(* IEC 61131-3 sources: daoli-st-library/DL_Base (part 13) *)

(* ---- FB_DL_InterlockMatrix.st ---- *)
(*==============================================================================
 * 组件名称 (Component)  : FB_DL_InterlockMatrix
 * 所属子库 (Sublibrary) : DL_Base
 * 当前版本 (Version)    : 1.0.1
 * 兼容性   (Platform)   : CODESYS 3.5 / TwinCAT 3 / 汇川 InoProShop / Machine Expert
 *                         仅依赖 Standard.library（R_TRIG / SHR / SHL），零厂商方言
 * 功能描述 (Function)   : 16 路安全联锁条件的汇总与首因（首出）追踪。
 *                         全部停机级条件满足才给出唯一一个运行许可位 bPermitToRun；
 *                         条件失效的瞬间锁存"第一个失效的通道号 + 完整位图 + 全局序号"，
 *                         复位后若条件仍未恢复，复位挂起而不清锁存。
 *                         解决两类现场顽疾：①停机后十条联锁同时报，维修工不知道先查哪条；
 *                         ②复位键一按就放行，根因被掩盖，第二天同一故障再来一次。
 *                         本块只回答"能不能开机"，"先看哪条报警"由报警管理组件负责。
 *
 * 【取反掩码真值表 / Invert-mask truth table（边界 B7）】
 *   raw  invert  →  有效值   现场含义
 *    0     0     →   0       常开触点未动作，条件不满足
 *    1     0     →   1       常开触点动作，条件满足
 *    0     1     →   1       常闭触点未断开（如未拍下的急停），条件满足
 *    1     1     →   0       常闭触点已断开（急停被拍下），条件不满足
 *   结论：常闭接线的急停、安全门、油压过低开关，必须把对应 invert 位置 1。
 *
 * 【失真与语义披露 / Distortion disclosure】
 *   1) 首因只在"停机级位图由 0 变非 0"的那一拍捕获。若两路在同一扫描周期内失效，
 *      扫描粒度内无法排序，此时取最低索引为代表值、置 bFirstOutSimult，并锁存整张位图；
 *      严禁在 HMI 上编造"谁先谁后"。
 *   2) 提示级失效不参与首因、不阻断许可，避免"料仓低"把停机首因挤掉。
 *   3) 上电首扫即锁存（不等沿）：冷启动时的首因可能只是"本来就断着"的条件，
 *      不代表本次停机原因，bLatchedAtStartup 用于区分这两种情形。
 *
 * 开源溯源 (Origin)     : 原创实现（参考 ISA-18.2 的首出方法论与西门子 LGF 位逻辑功能组的
 *                         参数分类，clean-room 编写，未复制任何源码）
 * 本文件内含       : TYPE  E_DL_InterlockState（配套枚举，归属 DL_Base）
 *                    FB    FB_DL_InterlockMatrix
 * 依赖     (Depends)    : 无 DL_ 内部依赖；Standard.library: R_TRIG / SHR / SHL
 * 红线自检 (Redline)    : R1 ✓ 零全局变量表与外部变量引用 ｜ R2 ✓ 零物理 IO 地址直写
 *                         R3 ✓ 纯 IEC 61131-3（位操作一律 SHR/SHL + AND/OR，无位访问方言）
 *                         R4 ✓ 配置非法即禁放行 + 复位挂起 + 序号饱和 + 索引钳位
 *                         R5 ✓ 全变量中英双语同行注释 ｜ R6 ✓ 五态 ENUM + CASE + ELSE 兜底
 *                         R7 ✓ 边沿实例主体最前部无条件刷新（本块仅一个实例）
 * 修订历史 (Revision)   :
 *   2026-11-14  v1.0.0  首版入库（Phase 1 收口批次 · R3）
 *   2026-11-16  v1.0.1  R13 机检 R39 修复：段 8 未使能覆盖原先把 eStateInt 无条件
 *                       改写为 eDisabled，而 eLatched / eFault 两态的复位沿消化
 *                       位于其后段 9 的 CASE 分支内——禁用期间按下的复位沿被整拍
 *                       吞掉，首因锁存与配置故障均需二次复位才清除。改为两个持有
 *                       复位沿的状态不被禁用覆盖，其余态行为不变
 *============================================================================*)

(*-----------------------------------------------------------------------------
 * 枚举: E_DL_InterlockState（归属 DL_Base，与 FB_DL_InterlockMatrix 同文件）
 * 含义: 联锁矩阵主状态。数值步长留空位便于后续插态而不破坏已有工程。
 *----------------------------------------------------------------------------*)
TYPE E_DL_InterlockState :
(
    eDisabled  := 0,     // 未使能：许可强制 FALSE，锁存内容保持 / Disabled, permit forced FALSE, latches kept
    eBlocked   := 10,    // 条件不满足：许可 FALSE，等待恢复 / Blocked, waiting for the conditions
    ePermitted := 20,    // 全部停机级条件满足，许可 TRUE / Permitted, all trip-class conditions OK
    eLatched   := 30,    // 首因已锁存，等待复位 / First-out latched, waiting for reset
    eFault     := 99     // 配置非法：无任何停机级通道，需改配置后复位 / Invalid configuration
);
END_TYPE

(*==============================================================================
 * 功能块: FB_DL_InterlockMatrix
 * 调用约定: 每个扫描周期无条件调用一次；abConditionOk 必须每拍整体刷新。
 * 无状态泄漏: 全部状态驻留于实例私有 VAR，零全局引用，可多机组并行实例化。
 *============================================================================*)
FUNCTION_BLOCK FB_DL_InterlockMatrix
VAR_INPUT
    abConditionOk : ARRAY[0..15] OF BOOL;     // 16 路原始条件，TRUE = 满足（上限 16 路）/ Raw conditions, TRUE = OK, max 16
    auInvertMask  : WORD := 16#0000;          // 取反掩码，bit=1 表示该路原始信号需取反 / Invert mask, bit=1 inverts that channel
    auTripMask    : WORD := 16#FFFF;          // 停机级掩码，bit=1 = 停机级，bit=0 = 提示级 / Trip-class mask, bit=1 is trip class
    bEnable       : BOOL := TRUE;             // 使能，FALSE 时许可 FALSE 且不清锁存 / Enable, FALSE forces permit down but keeps latches
    bReset        : BOOL;                     // 上升沿：清除首因锁存（条件未恢复则挂起）/ Rising edge: clear the first-out latch
END_VAR
VAR_OUTPUT
    bPermitToRun      : BOOL;                 // 运行许可（唯一放行信号）/ Run permit, the only release signal
    bFirstOutValid    : BOOL;                 // 首因有效 / First-out valid
    nFirstOutIndex    : INT;                  // 首因通道号 0..15，-1 = 无 / First-out channel 0..15, -1 = none
    uFirstOutMask     : WORD;                 // 首因位图（同拍多点时多 bit）/ First-out bitmap, multi-bit on simultaneous trips
    uFirstOutSeq      : UDINT;                // 首因发生的全局序号（单调递增）/ First-out global sequence, monotonic
    bFirstOutSimult   : BOOL;                 // 首因为同拍多点失效，扫描粒度内不可排序 / Simultaneous first-out, unorderable
    bLatchedAtStartup : BOOL;                 // 首因发生在上电首扫（冷启动即不满足）/ Latched during the first scan
    uTripActiveMask   : WORD;                 // 当前失效的停机级通道位图 / Currently failed trip channels
    uWarnActiveMask   : WORD;                 // 当前失效的提示级通道位图 / Currently failed warning channels
    bResetPending     : BOOL;                 // 复位挂起：已按复位但条件未恢复 / Reset pending, conditions not restored
    bError            : BOOL;                 // 故障标志（配置类锁存）/ Fault flag, configuration fault latched
    uErrorId          : UDINT;                // 故障码，0 = 无故障 / Error code, 0 = no error
    eState            : E_DL_InterlockState;  // 当前状态（供 HMI 诊断）/ Current state for HMI diagnosis
END_VAR
VAR
    fbTrigReset     : R_TRIG;                 // 复位上升沿检测实例 / Reset rising edge detector
    auEffOk         : ARRAY[0..15] OF BOOL;   // 取反后的有效条件（上限 16 路）/ Effective conditions after inversion, max 16
    uTripNow        : WORD;                   // 本拍失效的停机级位图 / Failed trip channels this scan
    uWarnNow        : WORD;                   // 本拍失效的提示级位图 / Failed warning channels this scan
    uPrevTripNow    : WORD;                   // 上一拍失效的停机级位图（判沿用）/ Previous trip bitmap, for edge detection
    uLatchMask      : WORD;                   // 锁存的首因位图 / Latched first-out bitmap
    uFirstOutSeqInt : UDINT;                  // 首因序号的内部副本 / Internal copy of the first-out sequence
    uBitMask        : WORD;                   // 单通道取位探针 / Single-channel bit probe
    nLatchIdx       : INT;                    // 锁存的首因通道号，-1 = 无 / Latched first-out index, -1 = none
    nNewLowest      : INT;                    // 本拍首个失效通道（最低索引）/ Lowest failed index this scan
    nBitCount       : INT;                    // 本拍失效通道总数 / Number of failed channels this scan
    nIdx            : INT;                    // 通道遍历索引 / Channel loop index
    uSeqCounter     : UDINT;                  // 全局序号计数器 / Global sequence counter
    eStateInt       : E_DL_InterlockState;    // 主状态机内部当前态 / Internal state of the main state machine
    bInv            : BOOL;                   // 该通道是否取反 / Whether this channel is inverted
    bConfigInvalid  : BOOL;                   // 本拍配置是否非法（无停机级通道）/ Configuration invalid this scan
    bConfigLatch    : BOOL;                   // 配置故障锁存 / Configuration fault latched
    bNewEvent       : BOOL;                   // 本拍出现新的停机级失效事件 / A new trip event started this scan
    bStartupScan    : BOOL := TRUE;           // 上电首扫标志 / First-scan flag
END_VAR
VAR CONSTANT
    DL_ILK_CHANNELS : INT  := 16;             // 通道数，必须等于数组维度 / Channel count, must match the array dimension
    DL_ILK_IDX_NONE : INT  := -1;             // 无效通道号哨兵 / No-channel sentinel
    DL_ILK_BIT0     : WORD := 16#0001;        // 最低位掩码 / Least significant bit mask
    DL_ILK_SEQ_MAX  : UDINT := 16#FFFF_FFFE;  // 序号饱和值 / Sequence saturation value
END_VAR

(*------------------------------------------------------------------------------
 * 段 1｜无条件刷新区（红线 R7）
 *      Unconditional refresh zone, placed at the very top of the body
 *-----------------------------------------------------------------------------*)
fbTrigReset(CLK := bReset);

(*------------------------------------------------------------------------------
 * 段 2｜上电首扫（边界 B2）：索引与位图必须显式置为哨兵值，不能依赖默认零
 *      First-scan init: the index must be forced to the sentinel, never left at zero
 *      0 号通道是合法的首因值，用 0 当"无首因"会让 HMI 永远显示 CH0 故障
 *-----------------------------------------------------------------------------*)
IF bStartupScan THEN
    nLatchIdx    := DL_ILK_IDX_NONE;
    uLatchMask   := 16#0000;
    uPrevTripNow := 16#0000;
    uSeqCounter  := 0;
    eStateInt    := E_DL_InterlockState.eBlocked;
END_IF

(*------------------------------------------------------------------------------
 * 段 3｜有效条件求值（边界 B7）：有效 = 原始 XOR 取反位
 *      Effective value = raw XOR invert, one pass over the 16 channels
 *      真值表见文件头；常闭接线的急停必须置 invert 位，否则"拍下急停"会被判为满足
 *      Normally-closed devices must set the invert bit, otherwise pressing the e-stop
 *      would read as a satisfied condition
 *-----------------------------------------------------------------------------*)
FOR nIdx := 0 TO (DL_ILK_CHANNELS - 1) DO
    uBitMask      := SHR(auInvertMask, nIdx) AND DL_ILK_BIT0;
    bInv          := (uBitMask <> 16#0000);
    auEffOk[nIdx] := abConditionOk[nIdx] XOR bInv;
END_FOR

(*------------------------------------------------------------------------------
 * 段 4｜分类汇总（边界 B6）：停机级进 uTripNow，提示级进 uWarnNow
 *      Classification: trip-class feeds the bitmap, warning-class only reports
 *      位操作一律 SHR/SHL 取位置位，禁止位访问方言，保证三平台同码
 *-----------------------------------------------------------------------------*)
uTripNow := 16#0000;
uWarnNow := 16#0000;

FOR nIdx := 0 TO (DL_ILK_CHANNELS - 1) DO
    IF NOT auEffOk[nIdx] THEN
        uBitMask := SHR(auTripMask, nIdx) AND DL_ILK_BIT0;
        IF uBitMask <> 16#0000 THEN
            uTripNow := uTripNow OR SHL(DL_ILK_BIT0, nIdx);
        ELSE
            uWarnNow := uWarnNow OR SHL(DL_ILK_BIT0, nIdx);
        END_IF
    END_IF
END_FOR

(*------------------------------------------------------------------------------
 * 段 5｜首因定位（边界 B3/B4）：求最低索引与失效总数
 *      First-out localisation: find the lowest failed index and the failed count
 *      同拍多路失效时无法排序，只能给代表值与位图，绝不编造先后
 *-----------------------------------------------------------------------------*)
nNewLowest := DL_ILK_IDX_NONE;
nBitCount  := 0;

FOR nIdx := 0 TO (DL_ILK_CHANNELS - 1) DO
    uBitMask := SHR(uTripNow, nIdx) AND DL_ILK_BIT0;
    IF uBitMask <> 16#0000 THEN
        nBitCount := nBitCount + 1;
        IF nNewLowest < 0 THEN
            nNewLowest := nIdx;
        END_IF
    END_IF
END_FOR

(*------------------------------------------------------------------------------
 * 段 6｜首因捕获：上电首扫特殊处理（边界 B2），其余按 0→非 0 的沿捕获
 *      First-out capture: special case on the first scan, edge-triggered afterwards
 *      锁存后不再被新故障覆盖——首因就是首因，覆盖等于把根因洗掉
 *      Once latched the value is never overwritten: the first cause stays the first cause
 *      首扫时 uPrevTripNow 已被置 0，因此"上电本来就不满足"同样走这条沿路径，
 *      只是序号从 1 开始并被标记为 bLatchedAtStartup
 *-----------------------------------------------------------------------------*)
bNewEvent := FALSE;

IF (uTripNow <> 16#0000) AND (uPrevTripNow = 16#0000) THEN
    bNewEvent := TRUE;
END_IF

IF bNewEvent THEN

    IF uSeqCounter < DL_ILK_SEQ_MAX THEN
        uSeqCounter := uSeqCounter + 1;
    ELSE
        uErrorId := 16#0001_0007;
    END_IF

    IF nLatchIdx < 0 THEN
        nLatchIdx         := nNewLowest;
        uLatchMask        := uTripNow;
        uFirstOutSeqInt   := uSeqCounter;
        bFirstOutSimult   := (nBitCount > 1);
        bLatchedAtStartup := bStartupScan;
    END_IF

END_IF

uPrevTripNow := uTripNow;

(*------------------------------------------------------------------------------
 * 段 7｜配置校验（边界 B1，fail-safe 第一原则）
 *      Configuration check: no trip-class channel means the permit can never be gated
 *      无任何停机级通道时若默认放行，等于把"没配置"当成"全部满足"，这是最危险的缺省
 *      Defaulting to permit when nothing is configured is the most dangerous default
 *-----------------------------------------------------------------------------*)
bConfigInvalid := (auTripMask = 16#0000);

IF bConfigInvalid THEN
    bConfigLatch := TRUE;
END_IF

IF bConfigLatch THEN
    uErrorId  := 16#0002_0004;
    eStateInt := E_DL_InterlockState.eFault;
END_IF

(*------------------------------------------------------------------------------
 * 段 8｜未使能处理：许可撤销、锁存保持（使能不是复位）
 *      Disabled: the permit drops but the latches survive, enabling is not resetting
 *      R39 纪律：复位沿只在发生的那一拍为真，其消化权归段 9 的 eLatched 与 eFault
 *      两个分支所有。本段若无条件把状态改写成 eDisabled，则禁用期间按下的复位沿
 *      在本拍即被抹掉（段 9 走 eDisabled 分支，两处复位判据都摸不到该沿），首因
 *      锁存与配置故障只能靠操作员补按第二次复位——故这两态不参与禁用覆盖。
 *      R39: the reset edge lives for exactly one scan and is consumed inside the CASE
 *      branches of eLatched and eFault, so the disable override must leave both
 *      states untouched; otherwise a reset pressed while disabled is lost and the
 *      first-out latch needs a second press. The other states keep the old behaviour.
 *-----------------------------------------------------------------------------*)
IF (eStateInt <> E_DL_InterlockState.eLatched)
AND (eStateInt <> E_DL_InterlockState.eFault)
AND (NOT bEnable) THEN
    eStateInt := E_DL_InterlockState.eDisabled;
END_IF

(*------------------------------------------------------------------------------
 * 段 9｜主状态机（红线 R6）：ENUM + CASE + ELSE 兜底
 *      Main state machine with the mandatory ELSE fallback
 *-----------------------------------------------------------------------------*)
CASE eStateInt OF

    E_DL_InterlockState.eDisabled:
        IF bEnable THEN
            IF bConfigLatch THEN
                eStateInt := E_DL_InterlockState.eFault;
            ELSE
                eStateInt := E_DL_InterlockState.eBlocked;
            END_IF
        END_IF

    E_DL_InterlockState.eBlocked:
        IF uTripNow <> 16#0000 THEN
            eStateInt := E_DL_InterlockState.eLatched;
        ELSE
            eStateInt := E_DL_InterlockState.ePermitted;
        END_IF

    E_DL_InterlockState.ePermitted:
        (* 任一停机级失效立即降级，许可在同一拍撤销（状态即许可） *)
        (* Any trip-class failure demotes at once, the permit drops in the same scan *)
        IF uTripNow <> 16#0000 THEN
            eStateInt := E_DL_InterlockState.eLatched;
        END_IF

    E_DL_InterlockState.eLatched:
        (* 边界 B5：条件未恢复时复位只挂起、不清锁存 *)
        (* Reset only pends while a trip condition is still present *)
        IF fbTrigReset.Q THEN
            IF uTripNow = 16#0000 THEN
                nLatchIdx         := DL_ILK_IDX_NONE;
                uLatchMask        := 16#0000;
                uFirstOutSeqInt   := 0;
                bFirstOutSimult   := FALSE;
                bLatchedAtStartup := FALSE;
                bResetPending     := FALSE;
                eStateInt         := E_DL_InterlockState.eBlocked;
            ELSE
                bResetPending := TRUE;
            END_IF
        END_IF

    E_DL_InterlockState.eFault:
        (* 配置故障：必须先把停机级掩码改对，再按复位退出 *)
        (* Configuration fault: fix the trip mask first, then reset *)
        IF fbTrigReset.Q AND (NOT bConfigInvalid) THEN
            bConfigLatch := FALSE;
            uErrorId     := 16#0000_0000;
            eStateInt    := E_DL_InterlockState.eBlocked;
        END_IF

    ELSE
        (* 非法状态拦截：不做隐式恢复，直接锁存上报 *)
        (* Illegal state interception: no implicit recovery, latch and report *)
        eStateInt := E_DL_InterlockState.eFault;
        uErrorId  := 16#0001_0005;

END_CASE;

(*------------------------------------------------------------------------------
 * 段 10｜输出单一出口（范式 P-05）
 *      Single output exit: the permit derives from the state exactly once
 *      分支内只改状态，许可位只在此处派生，"多处置位、漏撤一处"从结构上不可能
 *-----------------------------------------------------------------------------*)
bPermitToRun      := (eStateInt = E_DL_InterlockState.ePermitted) AND bEnable AND (NOT bConfigLatch);
bFirstOutValid    := (nLatchIdx >= 0);
nFirstOutIndex    := nLatchIdx;
uFirstOutMask     := uLatchMask;
uFirstOutSeq      := uFirstOutSeqInt;
uTripActiveMask   := uTripNow;
uWarnActiveMask   := uWarnNow;
bError            := (eStateInt = E_DL_InterlockState.eFault) OR bConfigLatch;
eState            := eStateInt;

(* 首扫标志在主体末尾撤销：段 6 需要它区分"冷启动即不满足"与"运行中失效" *)
(* The first-scan flag is cleared only here, stage 6 needs it for the cold-start case *)
bStartupScan := FALSE;
END_FUNCTION_BLOCK

(* ---- FB_DL_LastGoodValueHold.st ---- *)
(*
  ==================================================================
  组件名 Component  : FB_DL_LastGoodValueHold
  分类   Category   : DL_Base
  前缀   Naming     : FB_DL_ ｜ b/n/u/f/t/e 类型前缀制（R265）
  版本   Version    : 1.0.0
  功能   Purpose    : NE43 信号质量失效保持件：bSigOk=TRUE（质量好）时
                      透传 fInVal 并刷新保持载体；bSigOk=FALSE（NE43 超
                      量程/欠量程/断线诊断失效）时输出冻结为最后有效值
                      fLastGood，同时 tonStale 累计陈旧时长，超 tStaleMax
                      置信息码 01 与 bStale（输出仍保持最后有效值，不静
                      默）。失效时无历史有效值（首件语义）bValid=FALSE
                      并置信息码 03。tStaleMax ≤ 0 配置非法电平面码 02。
  来源   Source     : t2-8-ne43（NE43 欠量程/超量程诊断语义为公开行业
                      口径（NAMUR NE43），实现零源码复制）
  互引   Cross-ref  : FB_DL_AnalogOutFailsafe（同族失效安全件：其面向模
                      出通道失效替代，本件面向模拟量输入信号质量保持，
                      二者可级联——本件输出喂其输入）
  平台   Platform   : 纯 IEC 61131-3（TON/LREAL 四则/TIME 比较）
  依赖   Depends    : 仅 Standard.library（TON 属标准件）
  红线   Redline    : R1 零全局/VAR_EXTERNAL/R2 零 %I/%Q/R3 纯 IEC 标准
                      R4 输入非有限闸 + 配置闸显式 + TON 实例段 0 无条件
                      刷新/R5 全变量双语同行注释/R6 配置故障电平面无状
                      态机（CASE 不适用，头注说明）/R7 tonStale 无条件周
                      期调用/R8 阈值常量化
  契约   Contract   : 码 02 配置非法为电平面（当拍复判）：故障拍 bValid=
                      FALSE、fOut 冻结保持、bError=TRUE，恢复即恢复；
                      码 01/03 为信息级不置 bError。信号恢复（bSigOk 上
                      升）即透传刷新载体并清陈旧计时（TON 随 IN=FALSE
                      自清零，R188 自复位语义）。
  错误码 Codes      : 01【信息级】陈旧超限（保持时长超 tStaleMax，输出
                      仍为最后有效值）
                      02【故障级·电平面】tStaleMax ≤ T#0MS 配置非法
                      03【信息级】失效且无保持载体（从未收到有效值，
                      fOut 冻结 0）
  码位反证 Note     : 01/02/03 分立依据（R90）：01 在时效面（载体存在但
                      老化）、02 在配置面、03 在载体面（从未有过）可观测；
                      03 若并入 01，则「等一等会有值」与「永远不会有值」
                      不可区分，故必须分立；02 为故障级置 bError，与
                      01/03 信息级双通道可区分。
  验收   Acceptance : V1 质量好透传 → fOut=fInVal，bValid ｜ V2 失效 →
                      fOut 冻结最后值，bStale=FALSE（未超限）｜ V3 失效
                      超 tStaleMax → 码 01 + bStale ｜ V4 tStaleMax=0 →
                      码 02（电平面）｜ V5 上电即失效 → 码 03，bValid=
                      FALSE ｜ V6 恢复 → 透传 + 陈旧清零
  变更   Revision   : 2026-11-22  v1.0.0  R67 首版（编码阶段批 3 序 3）
  ==================================================================
*)
FUNCTION_BLOCK FB_DL_LastGoodValueHold
VAR_INPUT
    fInVal    : LREAL := 0.0;      // 输入测量值 [工程单位] / the input measured value
    bSigOk    : BOOL := FALSE;     // 信号质量好（NE43 诊断有效）[-] / the signal quality ok flag
    tStaleMax : TIME := T#60S;     // 陈旧时长上限 [ms]，须 > 0 / the staleness limit, must be positive
END_VAR
VAR_OUTPUT
    fOut     : LREAL := 0.0;       // 保持输出（最后有效值或透传）[工程单位] / the hold output
    bStale   : BOOL := FALSE;      // 陈旧超限指示（码 01 同源）[-] / the stale limit indicator
    bValid   : BOOL := FALSE;      // 输出可用标志（有有效载体且配置合法）[-] / the output usability flag
    bError   : BOOL := FALSE;      // 配置故障标志（电平面，恢复即清，R45 配对）/ the configuration fault flag
    uErrorId : UDINT := 16#0000_0000; // 错误码，0=正常，01/02/03 见头注 [码] / the error code [code]
END_VAR
VAR
    tonStale   : TON;              // 陈旧计时实例，段 0 无条件刷新 / the staleness timer instance refreshed unconditionally
    _fLastGood : LREAL := 0.0;     // 最后有效值保持载体 [工程单位] / the last good value hold carrier
    _bHasLast  : BOOL := FALSE;    // 保持载体是否存在（首件判据）[-] / the carrier existence flag
    _bCfgOk    : BOOL := FALSE;    // 本拍配置有效性 [-] / the per scan configuration validity
    _bSigFin   : BOOL := FALSE;    // 本拍输入有限性 [-] / the per scan input finiteness
END_VAR
VAR CONSTANT
    LGV_FIN_MAX  : LREAL := 1.7976931348623157E308; // LREAL 有限上限 / the finite LREAL limit
    LGV_ERR_NONE : UDINT := 16#0000_0000;           // 无错误 [码] / no error [code]
    LGV_ERR_STALE: UDINT := 16#0000_0001;           // 码 01：陈旧超限（信息级）/ code 01, stale limit, info level
    LGV_ERR_CFG  : UDINT := 16#0000_0002;           // 码 02：配置非法 / code 02, illegal configuration
    LGV_ERR_NOVAL: UDINT := 16#0000_0003;           // 码 03：无保持载体（信息级）/ code 03, no carrier, info level
END_VAR

(*------------------------------------------------------------------------------
 * 段 0｜定时器无条件刷新区（红线 R7）：严禁移入 IF / CASE
 *      The timer instance refreshes unconditionally, never inside a branch
 *-----------------------------------------------------------------------------*)
tonStale(IN := (NOT bSigOk) AND _bHasLast, PT := tStaleMax);  // 陈旧计时（失效且有载体才计时；恢复随 IN=FALSE 自清零，R188）/ the staleness timing, self clearing on recovery

(*------------------------------------------------------------------------------
 * 段 1｜错误码本拍预置 / segment 1, the error code per scan preset
 *-----------------------------------------------------------------------------*)
uErrorId := LGV_ERR_NONE;      // 预置无错误 / preset no error
bStale := FALSE;               // 陈旧指示预清（码 01 同源重算）/ preset the stale indicator

(*------------------------------------------------------------------------------
 * 段 2｜配置闸（电平面，当拍复判，码 02）+ 输入有限性闸
 *      The configuration gate and the input finiteness gate
 *-----------------------------------------------------------------------------*)
_bCfgOk := (tStaleMax > T#0MS);  // 配置闸（TIME 直接比较，三平台一致）/ the configuration gate
_bSigFin := (fInVal = fInVal) AND (ABS(fInVal) <= LGV_FIN_MAX);  // 输入非有限闸（NaN 自反判 + Inf 兜底）/ the input finite gate
IF NOT _bCfgOk THEN
    bError := TRUE;              // 故障标志（R45 配对）/ the fault flag
    uErrorId := LGV_ERR_CFG;     // 码 02 / code 02
    bValid := FALSE;             // 配置非法不出数 / no output on illegal configuration
    RETURN;                      // fOut 冻结保持（头注契约）/ the output frozen
ELSE
    bError := FALSE;             // 配置恢复即清（电平面契约）/ cleared when the configuration recovers
END_IF

(*------------------------------------------------------------------------------
 * 段 3｜质量好相：透传刷新载体（含非有限拒收，码 03 语义延用）
 *      The good quality phase, pass through and refresh the carrier
 *-----------------------------------------------------------------------------*)
IF bSigOk AND _bSigFin THEN
    _fLastGood := fInVal;        // 载体刷新 / refresh the carrier
    _bHasLast := TRUE;           // 载体存在 / the carrier exists
END_IF

(*------------------------------------------------------------------------------
 * 段 4｜失效相与出口映射：透传或保持，码 01/03 信息级
 *      The failed phase and the outlet mapping, the info codes
 *-----------------------------------------------------------------------------*)
IF bSigOk AND _bSigFin THEN
    fOut := fInVal;              // 透传 / pass through
ELSIF _bHasLast THEN
    fOut := _fLastGood;          // 保持最后有效值（锁存载体，非实时镜像混用）/ hold the last good value, the carrier not a live mirror
ELSE
    fOut := 0.0;                 // 无载体冻结 0（头注契约）/ frozen zero without a carrier
END_IF
IF (NOT bSigOk) OR (NOT _bSigFin) THEN
    IF NOT _bHasLast THEN
        uErrorId := LGV_ERR_NOVAL;  // 码 03：失效且从未有载体（信息级）/ code 03, no carrier, info level
        bValid := FALSE;            // 无值可保 / nothing to hold
    ELSE
        IF tonStale.Q THEN
            uErrorId := LGV_ERR_STALE;  // 码 01：陈旧超限（信息级，不置 bError）/ code 01, stale, info level
            bStale := TRUE;             // 陈旧指示（与码 01 同源，R191 名实双出口）/ the stale indicator
        END_IF
        bValid := TRUE;             // 有载体即可用（保持值有效语义）/ usable with a carrier
    END_IF
ELSE
    bValid := TRUE;                 // 质量好透传可用 / usable while passing through
END_IF
END_FUNCTION_BLOCK

(* ---- FB_DL_LongPressButton.st ---- *)
(*
  ==================================================================
  组件名 Component  : FB_DL_LongPressButton
  分类   Category   : DL_Base
  前缀   Naming     : FB_DL_ ｜ b/n/u/f/t/e/st 类型前缀制（R265）
  复杂度 Complexity  : 中
  版本   Version    : 1.0.0
  功能   Purpose    : 单按钮短按/长按/超长按三档时序分档（三窗 TON 阈值单拍分档）。
  来源   Source     : self-std（IEC 人机交互时序语义自研）
  平台   Platform   : 纯 IEC 61131-3（Standard.library: TON / R_TRIG / F_TRIG），无私有库
  分工声明 Split     : 与 FB_DL_ToggleButtonBank（模式解算属主）分工——后者做
                      按压次数模式解算；本件做单按钮按持续时长的三档分档
                      （R216 双向互引）。
  作者   Author     : 道莅代码库 · PLC 编程专家（R61）
  归属 Ownership     : 本件无 TYPE 声明；引用件类型全部 IEC 标准原生。
  ------------------------------------------------------------------
  边界 Boundary     :
                      一 三档窗组态闸（R239）：tShort < tLong < tXLong 且三者 > 0，
                         违反判组态非法故障码并冻结分档输出（锁存至复位沿）；
                      二 三窗职责与配比约束（R100）：tonShort < tonLong < tonXLong
                         由组态闸结构性保证；长按/超长按在按压持续中经阈值沿
                         单拍分档，短按在释放沿回判；
                      三 TON / R_TRIG / F_TRIG 全部段 0 无条件周期刷新（禁入分支）；
                      四 三档脉冲为单拍输出，段 1 统一预置 FALSE、分支只写 TRUE
                         （R256），内部 _b* 两段式映射（R187）；
                      五 故障态语义为「冻结保持全假输出」（R191 声明行）；
                      六 故障解除路径：复位沿清锁存（bReset 恒可达，R152 自证）；
                      七 无全局、无外部变量、无物理地址。
  错误码   Codes    :
    16#0001_0640【故障级】三档窗组态非法（tShort < tLong < tXLong 违反或 ≤0），锁存至复位沿
  验收   Acceptance :
    算法已证（脚本）：未跑 ｜ 编译器已证（三平台）：未跑
    V1 按下 200ms 释放（tShort=100/tLong=800/tXLong=2000）→ bShortPress 单拍
    V2 按住 1s → 长按阈值拍 bLongPress 单拍；V3 按住 2.5s → bXLongPress 单拍
    V4 tShort = tLong → 码 0640、三脉冲恒假、锁存待复位
  修订记录 Revision  :
    2026-11-21  v1.0.0  R61 首版（批 2 · 序号 8）
  ==================================================================
*)
FUNCTION_BLOCK FB_DL_LongPressButton
VAR_INPUT
    bBtn   : BOOL := FALSE; // 按钮输入电平 [-] / the button input level
    bReset : BOOL := FALSE; // 故障复位电平，上升沿清锁存 [-] / the fault reset level
    tShort : TIME := T#100MS; // 短按下限阈值 [毫秒]，须 < tLong / the short press lower threshold
    tLong  : TIME := T#800MS; // 长按阈值 [毫秒]，须 < tXLong / the long press threshold
    tXLong : TIME := T#2S;    // 超长按阈值 [毫秒] / the extra long press threshold
END_VAR
VAR_OUTPUT
    bShortPress : BOOL := FALSE; // 短按单拍脉冲（释放沿回判）[-] / the short press one shot
    bLongPress  : BOOL := FALSE; // 长按单拍脉冲（tLong 阈值沿）[-] / the long press one shot
    bXLongPress : BOOL := FALSE; // 超长按单拍脉冲（tXLong 阈值沿）[-] / the extra long press one shot
    bFaulted    : BOOL := FALSE; // 组态故障锁存指示 [-] / the latched configuration fault indicator
    eErr        : UDINT := 16#0000_0000; // 错误码，0 = 正常 / the error code, zero is ok
    bError      : BOOL := FALSE; // 故障锁存位（与锁存同源，R191）/ the fault bit from the same latch
END_VAR
VAR
    _bInit      : BOOL := FALSE; // 首拍初始化标志（R310）/ the first scan flag
    _bFault     : BOOL := FALSE; // 组态故障锁存副本（仅复位沿清除）/ the fault latch copy
    _bShort     : BOOL := FALSE; // 短拍内部位，段 1 预清段 5 映射 / the internal short bit
    _bLong      : BOOL := FALSE; // 长拍内部位 / the internal long bit
    _bXLong     : BOOL := FALSE; // 超长拍内部位 / the internal extra long bit
    _bLongFired : BOOL := FALSE; // 长按已发标记（释放沿判短按排除用，按压期间保持）/ the long fired flag held during the press
    _bXFired    : BOOL := FALSE; // 超长按已发标记 / the extra long fired flag
    _bCfgBad    : BOOL := FALSE; // 组态非法标记（逐拍重算）/ the configuration fault flag recomputed
    rtBtn       : R_TRIG;  // 按钮按下沿实例，段 0 无条件刷新 / the press edge instance
    ftBtn       : F_TRIG;  // 按钮释放沿实例，段 0 无条件刷新 / the release edge instance
    rtReset     : R_TRIG;  // 复位沿实例，段 0 无条件刷新 / the reset edge instance
    rtLongQ     : R_TRIG;  // 长窗到时沿实例，段 0 无条件刷新 / the long window expiry edge instance
    rtXLongQ    : R_TRIG;  // 超长窗到时沿实例，段 0 无条件刷新 / the extra long expiry edge instance
    tonShort    : TON;     // 短窗计时，段 0 无条件刷新 / the short window timer
    tonLong     : TON;     // 长窗计时 / the long window timer
    tonXLong    : TON;     // 超长窗计时 / the extra long window timer
END_VAR

// 段 0｜定时器与沿检测无条件周期刷新（禁入分支，R7）/ segment 0, the unconditional refresh
rtBtn(CLK := bBtn); // 按下沿 / the press edge
ftBtn(CLK := bBtn); // 释放沿 / the release edge
rtReset(CLK := bReset); // 复位沿 / the reset edge
tonShort(IN := bBtn, PT := tShort); // 短窗计时（按压电平驱动）/ the short window timing
tonLong(IN := bBtn, PT := tLong); // 长窗计时 / the long window timing
tonXLong(IN := bBtn, PT := tXLong); // 超长窗计时 / the extra long window timing
rtLongQ(CLK := tonLong.Q); // 长窗到时沿 / the long expiry edge
rtXLongQ(CLK := tonXLong.Q); // 超长窗到时沿 / the extra long expiry edge

// 段 1｜首拍初始化与单拍标志预清（仅单拍标志入清单，FB32-1；R256）/ segment 1, the first scan init and the one shot preset
IF NOT _bInit THEN // 首拍一拍 / the first scan
    _bInit := TRUE; // 置首拍标志 / raise the first scan flag
    _bFault := FALSE; // 故障锁存显式清零 / clear the fault latch explicitly
    _bLongFired := FALSE; // 长发标记显式清零 / clear the long fired flag explicitly
    _bXFired := FALSE; // 超长发标记显式清零 / clear the extra long fired flag explicitly
END_IF
IF rtReset.Q THEN // 复位沿：清故障锁存（解除路径：复位沿恒可达，R152 自证）/ the reset edge clears the latch
    _bFault := FALSE; // 清锁存 / clear the latch
END_IF
_bShort := FALSE; // 短拍预清零 / preset the short bit false
_bLong := FALSE; // 长拍预清零 / preset the long bit false
_bXLong := FALSE; // 超长拍预清零 / preset the extra long bit false
_bCfgBad := FALSE; // 组态标记预清零 / preset the configuration flag false

// 段 2｜组态域闸（三窗严格递增 + 正值，R239，边界一）/ segment 2, the configuration gate
IF (tShort <= T#0S) OR (tLong <= tShort) OR (tXLong <= tLong) THEN // 递增配比违反或非正 / the monotone ratio violated
    _bCfgBad := TRUE; // 置组态非法标记 / raise the configuration flag
    _bFault := TRUE; // 锁存故障（段 5 出口回放）/ latch the fault
END_IF

// 段 3｜按压中阈值沿分档（故障冻结，边界五；沿只在合法态消费）/ segment 3, the threshold edges during the press
IF (NOT _bFault) AND bBtn THEN // 合法态且按压中 / legal and pressed
    IF rtLongQ.Q AND (NOT _bLongFired) AND (NOT _bXFired) THEN // 长窗到时沿首现 / the long expiry edge first seen
        _bLong := TRUE; // 置长拍 / raise the long bit
        _bLongFired := TRUE; // 锁长发标记（释放沿判短按排除）/ latch the long fired flag
    END_IF
    IF rtXLongQ.Q AND (NOT _bXFired) THEN // 超长窗到时沿首现 / the extra long expiry edge first seen
        _bXLong := TRUE; // 置超长拍 / raise the extra long bit
        _bXFired := TRUE; // 锁超长发标记 / latch the extra long fired flag
    END_IF
END_IF

// 段 4｜释放沿回判短按（短按 = 释放时短窗已到而长按未发，边界二）/ segment 4, the release edge judges the short press
IF ftBtn.Q AND (NOT _bFault) THEN // 合法态释放沿 / a legal release edge
    IF tonShort.Q AND (NOT _bLongFired) AND (NOT _bXFired) THEN // 短窗已到且未触发高档 / the short window met with no higher grade fired
        _bShort := TRUE; // 置短拍 / raise the short bit
    END_IF
    _bLongFired := FALSE; // 释放清长发标记（下一按压新起点）/ clear the long fired flag at the release
    _bXFired := FALSE; // 释放清超长发标记 / clear the extra long fired flag
END_IF

// 段 5｜统一出口（内部副本单点映射；故障冻结全假，R191）/ segment 5, the unified outlet with the frozen fault
bShortPress := _bShort AND (NOT _bFault); // 短拍出口 / the short outlet
bLongPress := _bLong AND (NOT _bFault); // 长拍出口 / the long outlet
bXLongPress := _bXLong AND (NOT _bFault); // 超长拍出口 / the extra long outlet
bFaulted := _bFault; // 故障指示出口 / the fault indicator outlet
bError := _bFault; // 故障位出口（与锁存同源，R191）/ the fault bit outlet
IF _bFault THEN // 故障锁存回放（R187）/ the latched fault replays
    eErr := 16#0001_0640; // 故障级：三档窗组态非法 / fault grade, the illegal window configuration
ELSE // 无故障 / no fault
    eErr := 16#0000_0000; // 正常 / ok
END_IF
END_FUNCTION_BLOCK

(* ---- FB_DL_ManualOverride.st ---- *)
(*
  道莅工业代码库 | DL_Base | FB_DL_ManualOverride
  版本: 1.0.0 | 日期: 2026-11-23 | 轮次: R75
  开源溯源: brOscatLib (github.com/brOscatLib) / MIT / 借鉴 MANUAL 覆写的语义，代码为 clean-room 重写
  功能: 手动强制覆写——覆写请求上升沿激活后输出切手动值，最长保持 tMaxHold
        （T#0S = 无限时）超时自动回落自动值；释放沿/禁止输入即时回落；
        激活单拍提示脉冲与超时回落信息码。
  兼容性: CODESYS 3.5 / TwinCAT 3 / 汇川 InoProShop；仅依赖标准 TON / R_TRIG / SEL，零厂商私有库
  接口: 输入 bOverrideReq（沿）/bRelease（沿）/fAutoVal/fManualVal/tMaxHold/
        bInhibit/bReset；输出 bOverride/bOut/bActPulse/bTimedOut/eState/eInfo/nErrId。
  码表: 16#0001_04BC 信息级：覆写超时自动回落（锁存至复位沿）
        16#0001_04BD 信息级：覆写请求被禁止拒绝（当拍重算）
        16#0001_04BE 信息级：覆写中手动值非有限（输出保持最后有效值，当拍重算）
        码段说明：0001 段信息子带 04xx，槽位经全库实扫空闲。
  边界: ① 手动值 NaN 拒绝激活（待机相判码），覆写中手动值变 NaN → 输出保持
        最后有效值并置信息码（冻结语义不穿透坏值）；
        ② bInhibit 在覆写中即时回落自动值（禁止优先于覆写，安全侧）；
        ③ 超时判定仅当 tMaxHold > T#0S 生效（T#0S = 无限保持）；
        ④ TON/R_TRIG 段 0 无条件周期刷新；⑤ 本件全部事件均为信息级，无故障级码；
        ⑥ 零全局耦合。
  邻件比对: ToleranceWindow（单容差窗）与本件无语义交集；S04 E_DL_ControlModeSel
            为本件模式语义配套枚举（后续入库）。
  修订历史: 2026-11-23 v1.0.0 R75 首版（复杂件批 B3 · C11）
*)

TYPE E_DL_MovState :
(
    eIdle    := 0,   // 覆写未激活（输出自动值） | Override inactive, output auto value
    eActive  := 10   // 覆写激活（输出手动值） | Override active, output manual value
);
END_TYPE

TYPE E_DL_MovInfo :
(
    eNone      := 0,  // 无事件 | No event
    eTimeout   := 1,  // 超时自动回落（锁存至复位沿） | Timed out, auto fallback latched
    eInhibit   := 2,  // 请求被禁止拒绝（当拍重算） | Request rejected by inhibit
    eNonFinite := 3   // 手动值非有限（当拍重算，输出保持） | Manual value non-finite, output held
);
END_TYPE

FUNCTION_BLOCK FB_DL_ManualOverride
VAR_INPUT
    bOverrideReq : BOOL := FALSE;   // 覆写请求（上升沿激活）[-] | Override request, rising edge activates
    bRelease     : BOOL := FALSE;   // 释放请求（上升沿回落）[-] | Release request, rising edge falls back
    fAutoVal     : REAL := 0.0;     // 自动值 [工程单位] | Auto value
    fManualVal   : REAL := 0.0;     // 手动值（覆写目标）[工程单位] | Manual value, override target
    tMaxHold     : TIME := T#30S;   // 最长覆写保持，T#0S = 无限 | Max hold duration, T#0S = unlimited
    bInhibit     : BOOL := FALSE;   // 覆写禁止（电平，覆写中即时回落）[-] | Override inhibit level
    bReset       : BOOL := FALSE;   // 复位命令，上升沿清超时锁存 [-] | Reset command, rising edge
END_VAR
VAR_OUTPUT
    bOverride : BOOL;               // 覆写激活态 [-] | Override active state
    fOut      : REAL;               // 选择输出（自动/手动/保持值）[工程单位] | Selected output value
    bActPulse : BOOL;               // 激活单拍提示脉冲 [-] | Activation one-shot pulse
    bTimedOut : BOOL;               // 超时回落锁存标志 [-] | Timed-out latch flag
    eState    : E_DL_MovState;      // 状态出口 | State outlet
    eInfo     : E_DL_MovInfo;       // 事件成因出口 | Event cause outlet
    nErrId    : UDINT;              // 事件码，0 = 无事件 | Event code, 0 = none
END_VAR
VAR
    _eState    : E_DL_MovState := E_DL_MovState.eIdle;   // 内部状态（CASE 唯一写入目标） | Internal state
    _eInfo     : E_DL_MovInfo := E_DL_MovInfo.eNone;     // 事件成因锁存（超时级） | Latched event cause
    _bOverride : BOOL;          // 覆写激活锁存位 | Override active latch bit
    _bTimedOut : BOOL;          // 超时回落锁存位 | Timed-out latch bit
    _bHold     : BOOL;          // 输出保持当拍量（手动值非有限）[-] | Output hold this scan
    _fOutLast  : REAL := 0.0;   // 最后有效输出保持值 [工程单位] | Last valid output hold value
    _bNonFin   : BOOL;          // 手动值非有限当拍量 [-] | Manual value non-finite this scan
    _uInfo     : UDINT;         // 信息码每拍重算 | Info code per scan
    rtReq      : R_TRIG;        // 覆写请求沿实例，段 0 无条件刷新 | Override request edge instance
    rtRel      : R_TRIG;        // 释放沿实例，段 0 无条件刷新 | Release edge instance
    rtReset    : R_TRIG;        // 复位沿实例，段 0 无条件刷新 | Reset edge instance
    rtAct      : R_TRIG;        // 激活沿实例（单拍提示），段 0 无条件刷新 | Activation edge instance for one-shot
    tonHold    : TON;           // 覆写保持计时，段 0 无条件刷新 | Override hold timer
END_VAR

(* —— 段 0：当拍量派生 + 定时器与沿实例无条件周期刷新（R7 红线） —— *)
_bNonFin := (fManualVal <> fManualVal);                                     // 手动值 NaN 自反判 / Manual value NaN self-reflex check
rtReq(CLK := bOverrideReq);                                                 // 请求沿每拍必调 / Request edge every scan
rtRel(CLK := bRelease);                                                     // 释放沿每拍必调 / Release edge every scan
rtReset(CLK := bReset);                                                     // 复位沿每拍必调 / Reset edge every scan
rtAct(CLK := _bOverride);                                                   // 激活态沿（单拍提示用）每拍必调 / Activation edge for one-shot
tonHold(IN := (_eState = E_DL_MovState.eActive) AND (tMaxHold > T#0S), PT := tMaxHold);  // 保持计时，IN 挂激活 ∧ 有限时限 / Hold timer gated by active and finite limit

(* —— 段 1：复位沿清超时锁存 —— *)
IF rtReset.Q THEN
    _bTimedOut := FALSE;                                                    // 清超时锁存位 / Clear timed-out latch
    _eInfo := E_DL_MovInfo.eNone;                                           // 清成因锁存 / Clear latched cause
END_IF

(* —— 段 2：状态机（ENUM + CASE，ELSE 兜底） —— *)
CASE _eState OF

E_DL_MovState.eIdle:
    IF rtReq.Q AND bInhibit THEN
        _uInfo := 16#0001_04BD;                                             // 信息级：请求被禁止拒绝 / Info: request rejected by inhibit
    ELSIF rtReq.Q AND _bNonFin THEN
        _uInfo := 16#0001_04BE;                                             // 信息级：手动值非有限拒绝激活 / Info: non-finite manual refused
    ELSIF rtReq.Q THEN
        _bOverride := TRUE;                                                 // 激活覆写锁存 / Activate override latch
        _eState := E_DL_MovState.eActive;                                   // 进入激活相 / Enter active phase
    END_IF

E_DL_MovState.eActive:
    IF rtRel.Q THEN
        _bOverride := FALSE;                                                // 释放沿回落 / Release edge falls back
        _eState := E_DL_MovState.eIdle;
    ELSIF bInhibit THEN
        _bOverride := FALSE;                                                // 禁止输入即时回落（安全侧优先，边界②）/ Inhibit forces fallback
        _eState := E_DL_MovState.eIdle;
    ELSIF tonHold.Q THEN
        _bOverride := FALSE;                                                // 超时回落 / Timed out, fall back
        _bTimedOut := TRUE;                                                 // 超时锁存（复位沿清）/ Latch timeout
        _eInfo := E_DL_MovInfo.eTimeout;                                    // 归因超时 / Cause: timeout
        _eState := E_DL_MovState.eIdle;
    END_IF

ELSE
    _eState := E_DL_MovState.eIdle;                                         // 非法状态兜底（R6，回落安全侧）/ Illegal state fallback to safe side
    _bOverride := FALSE;                                                    // 非法态覆写强制撤 / Override forced off

END_CASE

(* —— 段 3：出口单点映射（名实同源；选择 + 保持 + 锁存码回放） —— *)
IF _bOverride AND _bNonFin THEN
    _bHold := TRUE;                                                         // 覆写中手动值变坏：保持当拍置位（边界①）/ Manual went bad while active, hold
    _uInfo := 16#0001_04BE;                                                 // 信息级：手动值非有限 / Info: manual non-finite
ELSE
    _bHold := FALSE;                                                        // 正常拍不保持 / No hold on normal scan
END_IF
IF (NOT _bHold) AND (NOT (_bOverride AND _bNonFin)) THEN
    _fOutLast := fManualVal;                                                // 有效拍刷新保持值（手动值载体）/ Refresh hold value on valid manual
END_IF
bOverride := _bOverride;                                                    // 覆写态镜像 / Override mirror
IF _bOverride AND _bNonFin THEN
    fOut := _fOutLast;                                                      // 坏值拍输出保持值（冻结语义）/ Bad-value scan outputs held value
ELSIF _bOverride THEN
    fOut := fManualVal;                                                     // 覆写输出手动值 / Override outputs manual value
ELSE
    fOut := fAutoVal;                                                       // 未覆写输出自动值 / Idle outputs auto value
END_IF
bActPulse := rtAct.Q;                                                       // 激活单拍提示（R_TRIG 单拍化） / Activation one-shot
bTimedOut := _bTimedOut;                                                    // 超时锁存镜像 / Timeout latch mirror
eState := _eState;                                                          // 状态出口 / State outlet
eInfo := _eInfo;                                                            // 成因出口 / Cause outlet
IF _bTimedOut THEN
    nErrId := 16#0001_04BC;                                                 // 超时回落锁存码回放（最高优先）/ Replay timeout code
ELSIF _uInfo <> 16#0000_0000 THEN
    nErrId := _uInfo;                                                       // 当拍信息码 / Per-scan info code
ELSE
    nErrId := 16#0000_0000;                                                 // 无事件 / No event
END_IF

END_FUNCTION_BLOCK

(* ---- FB_DL_MinOnOffGuard.st ---- *)
(*
    组件名称 : FB_DL_MinOnOffGuard
    所属子库 : DL_Base
    当前版本 : 1.0.0
    兼 容 性 : CODESYS V3.5+ / TwinCAT 3 / 汇川 InoProShop；仅依赖 Standard.library
    功能描述 : 最短运行 / 最短停止双守卫，防压缩机、热泵、泵轮值与冷水机组频繁启停的公共原子。
              取舍 ①：用「输出实际在 TRUE 期间的累计时长」判最短运行，而不是「进入某状态后重新计时」——
              若定时器只在 eStarting 与 eHolding 里跑，请求在 eRunning 撤掉后会重新起算整段 tMinOn，
              实际运行时长翻倍，压缩机照样被拖坏。本件把 eRunning 一并纳入定时器 IN，
              于是 fbMinOn.Q 的语义严格等于「输出已持续 TRUE 达到 tMinOn」。
              取舍 ②：eIdle 的启动条件只看 bReq，不再二次判 fbMinOff.Q —— 若 eIdle 还要等最短停止完成位，
              而该定时器只在 eCooldown 里通电，则 Q 在 eIdle 恒为 FALSE，状态机将永远起不来（本件修正了这个死锁形态）。
              最短停止由「必须走完 eCooldown 才回 eIdle」保证，语义不减。
              取舍 ③：参数非法不停机 —— 守卫时间填成负值属于参数错误，钳零后继续跑并发故障码；
              让一条产线因为一个 HMI 输入框的负号而停机，代价远大于收益。
              取舍 ④：bEnable = FALSE 走安全侧 —— 立即输出 FALSE 并回 eIdle，忽略最短运行；
              安全优先于设备寿命，两者冲突时永远选安全。
    开源溯源 : 原创实现（T0-2 变体线）。ROADMAP 中「防频繁启停」四条待办的公共原子，无外部源码参考，；本件为 IEC 61131-3 标准语义的道莅防御性实现（原创实现，零外部源码复制）。
              状态机、码位、钳位策略 100% 自有。
    本文件内含 : FUNCTION_BLOCK FB_DL_MinOnOffGuard
                 同文件 TYPE E_DL_MinOnOffState（归属本子库，全库唯一）
    依 赖 : 无 DL_ 内部依赖；Standard.library: TON / R_TRIG
    红线自检 : R1 ✓ 零全局变量与外部变量 ｜ R2 ✓ 零物理 IO 地址
              R3 ✓ 纯 IEC 61131-3 ｜ R4 ✓ 参数钳位 + 非法时间闸 + 非法状态 ELSE 兜底 + 复位沿优先
              R5 ✓ 全变量中英双语同行注释 ｜ R6 ✓ ENUM + CASE + ELSE 兜底（非法状态落 039A 并回安全态）
              R7 ✓ TON / R_TRIG 实例在主体最前部无条件刷新，位于任何 IF 与 CASE 之外
              R8 ✓ 时间上限、零时长、错误码全常量化
    错误码   : 16#0001_0452 [信息级] 时间参数超 24h 已钳上限，bError = FALSE
               16#0001_0453 [信息级] 停机请求被最短运行推迟（进入 eHolding），bError = FALSE
               16#0001_0399 [故障级] 时间参数为负已钳零，不停机，bError = TRUE
               16#0001_039A [故障级] 非法状态（枚举被改写），强制回 eFault 且 bOut = FALSE
               16#0001_039B [故障级] 预留禁用（不得挪用）
    码位总账 : 16#0001_0452 用 / 16#0001_0453 用 ｜ 16#0001_0399 用 / 16#0001_039A 用 / 16#0001_039B 预留
              说明：「启动请求被最短停止阻延」不设独立码 —— 该场景由 eState = eCooldown、bHoldOff 与 tRemaining
              三个输出直接可观测，加强加码属凑槽（R90）。
    遗留假设 : ① TIME 比较与减法按 32 位有符号毫秒口径，加减不越 24h 上限（已由钳位保证），
              故无 TIME 回绕路径；该推导未在三平台逐一实测。
              ② bReset 只在 eFault 内被消费（复位沿实例仍在主体最前部刷新），保证复位沿不被 CASE 前置写吞掉。
    修订历史 :
        2026-11-16  v1.0.0  首版，R21 批次 4 入库
*)

(*-----------------------------------------------------------------------------
 * 枚举: E_DL_MinOnOffState（归属本功能块，与其同文件发布，全库唯一）
 * 含义: 双守卫状态机的六个状态，成员值写死便于工程持久化与在线诊断
 *----------------------------------------------------------------------------*)
TYPE E_DL_MinOnOffState :
(
    eIdle     := 0,     // 空闲：输出 FALSE，最短停止已满，可随时启动 / idle, output low and the minimum off time is satisfied
    eStarting := 10,    // 启动中：输出 TRUE，最短运行计时中 / starting, output high and the minimum on time is counting
    eRunning  := 20,    // 运行中：输出 TRUE，最短运行已满 / running, the minimum on time is satisfied
    eHolding  := 30,    // 保持中：请求已撤但最短运行未满，强制输出 TRUE / holding, the request is gone but the minimum on time is not yet met
    eCooldown := 40,    // 冷却中：输出 FALSE，最短停止计时中 / cooling down, output low and the minimum off time is counting
    eFault    := 99     // 故障锁定：输出 FALSE，需 bReset 上升沿退出 / fault latched, cleared by the rising edge of bReset
);
END_TYPE

FUNCTION_BLOCK FB_DL_MinOnOffGuard
VAR_INPUT
    bEnable         : BOOL := TRUE;      // 使能，FALSE 立即回安全态并忽略最短运行 / enable, FALSE forces the safe state and ignores the minimum on time
    bReq            : BOOL;              // 上层运行请求，TRUE 表示希望设备运行 / run request from the upper layer
    tMinOn          : TIME := T#10S;     // 最短运行时间，负值钳零、超 24h 钳上限 [ms] / minimum on time, clamped at both ends [ms]
    tMinOff         : TIME := T#10S;     // 最短停止时间，负值钳零、超 24h 钳上限 [ms] / minimum off time, clamped at both ends [ms]
    bReset          : BOOL;              // 上升沿清故障并回空闲 / rising edge clears the fault and returns to idle
END_VAR
VAR_OUTPUT
    bOut            : BOOL;              // 实际输出，最终的启停指令 / effective output, the final run command
    bHoldOn         : BOOL;              // TRUE = 正在强制延长运行（停机请求被推迟）/ TRUE while the run time is being extended
    bHoldOff        : BOOL;              // TRUE = 正在强制延长停止（启动请求被阻延）/ TRUE while the stop time is being extended
    tRemaining      : TIME;              // 当前守卫的剩余时间，无守卫时为 0 [ms] / remaining guard time, zero when no guard is active [ms]
    eState          : E_DL_MinOnOffState;   // 状态机当前状态 / current state machine state
    eErr            : UDINT;             // 错误码，0=正常；16#0001_04XX 信息级 / 16#0001_03XX 故障级 / error id, 0=ok
    bError          : BOOL;              // 故障级标志，eErr 落 16#0001_03XX 时为 TRUE / fault flag, TRUE on fault-level eErr
END_VAR
VAR
    fbMinOn         : TON;               // 最短运行计时器，主体最前部无条件刷新 / minimum on timer, refreshed unconditionally at the top
    fbMinOff        : TON;               // 最短停止计时器，主体最前部无条件刷新 / minimum off timer, refreshed unconditionally at the top
    rtReset         : R_TRIG;            // 复位上升沿，主体最前部无条件刷新 / reset rising edge, refreshed unconditionally at the top
    tMinOnEff       : TIME;              // 钳位后的最短运行时间 [ms] / clamped minimum on time [ms]
    tMinOffEff      : TIME;              // 钳位后的最短停止时间 [ms] / clamped minimum off time [ms]
END_VAR
VAR CONSTANT
    DL_MIN_ONOFF_MAX    : TIME := T#24H;               // 守卫时间上限，超此值无工程意义 [ms] / guard time upper bound [ms]
    DL_TIME_ZERO        : TIME := T#0S;                // 零时长哨兵 [ms] / zero duration sentinel [ms]
    DL_ERR_NONE         : UDINT := 16#0000_0000;       // 无故障 / no error
END_VAR

// 段 0｜错误状态预置（四段式第一段）/ segment 0, preset the error state
eErr   := DL_ERR_NONE;                  // 预置无错误 / preset no error
bError := FALSE;                        // 预置无故障 / preset no fault

// 段 1｜参数预处理：本段无任何定时器调用，故可置于定时器刷新之前，保证钳位当拍生效 / segment 1, pure parameter preprocessing
tMinOnEff  := tMinOn;                   // 先按输入占位 / start from the input
tMinOffEff := tMinOff;                  // 先按输入占位 / start from the input
IF tMinOnEff < DL_TIME_ZERO THEN
    tMinOnEff := DL_TIME_ZERO;          // 负值钳零，不停机 / clamp to zero, the machine keeps running
    eErr      := 16#0001_0399;          // 时间参数为负（故障级）/ negative time parameter, fault level
    bError    := TRUE;                  // 置故障标志 / raise the fault flag
END_IF
IF tMinOffEff < DL_TIME_ZERO THEN
    tMinOffEff := DL_TIME_ZERO;         // 负值钳零 / clamp to zero
    eErr       := 16#0001_0399;         // 同一语义，同一码 / one semantic, one code
    bError     := TRUE;                 // 置故障标志 / raise the fault flag
END_IF
IF tMinOnEff > DL_MIN_ONOFF_MAX THEN
    tMinOnEff := DL_MIN_ONOFF_MAX;      // 超上限钳位 / clamp above the bound
    IF eErr = DL_ERR_NONE THEN
        eErr := 16#0001_0452;           // 参数超上限已钳位（信息级）/ parameter clamped, info level
    END_IF
END_IF
IF tMinOffEff > DL_MIN_ONOFF_MAX THEN
    tMinOffEff := DL_MIN_ONOFF_MAX;     // 超上限钳位 / clamp above the bound
    IF eErr = DL_ERR_NONE THEN
        eErr := 16#0001_0452;           // 参数超上限已钳位（信息级）/ parameter clamped, info level
    END_IF
END_IF

// 段 2｜定时器与边沿无条件刷新：位于任何 IF 与 CASE 之外（红线 R7）/ segment 2, unconditional timer refresh
fbMinOn ( IN := (eState = E_DL_MinOnOffState.eStarting) OR (eState = E_DL_MinOnOffState.eHolding) OR (eState = E_DL_MinOnOffState.eRunning),
          PT := tMinOnEff );
fbMinOff( IN := (eState = E_DL_MinOnOffState.eCooldown), PT := tMinOffEff );
rtReset ( CLK := bReset );

// 段 3｜失能走安全侧：唯一允许的 CASE 前置状态改写，条件由 bEnable 限定 / segment 3, the only pre-CASE write, guarded by the enable
IF NOT bEnable THEN
    eState := E_DL_MinOnOffState.eIdle;  // 立即回空闲，最短运行让位于安全 / back to idle at once, safety outranks machine life
END_IF

// 段 4｜状态机 / segment 4, state machine
CASE eState OF
    E_DL_MinOnOffState.eIdle :
        bOut := FALSE;                                          // 空闲输出低 / idle output is low
        IF bReq THEN
            eState := E_DL_MinOnOffState.eStarting;             // 有请求即启动，最短停止已在 eCooldown 走完 / start on request, the off time was already served
        END_IF

    E_DL_MinOnOffState.eStarting :
        bOut := TRUE;                                           // 启动中输出高 / output is high while starting
        IF fbMinOn.Q THEN
            eState := E_DL_MinOnOffState.eRunning;              // 最短运行已满 / the minimum on time is satisfied
        END_IF

    E_DL_MinOnOffState.eRunning :
        bOut := TRUE;                                           // 运行中输出高 / output is high while running
        IF NOT bReq THEN
            IF NOT fbMinOn.Q THEN
                IF eErr = DL_ERR_NONE THEN
                    eErr := 16#0001_0453;                       // 停机请求被最短运行推迟（信息级）/ the stop request is delayed by the minimum on time
                END_IF
            END_IF
            eState := E_DL_MinOnOffState.eHolding;              // 进入保持态，由定时器完成位决定何时真正停机 / enter holding, the timer decides
        END_IF

    E_DL_MinOnOffState.eHolding :
        bOut := TRUE;                                           // 保持中仍输出高 / output stays high while holding
        IF fbMinOn.Q THEN
            eState := E_DL_MinOnOffState.eCooldown;             // 最短运行补满，进入冷却 / the minimum on time is met, cool down
        END_IF

    E_DL_MinOnOffState.eCooldown :
        bOut := FALSE;                                          // 冷却输出低 / output is low while cooling down
        IF fbMinOff.Q THEN
            eState := E_DL_MinOnOffState.eIdle;                 // 最短停止已满 / the minimum off time is satisfied
        END_IF

    E_DL_MinOnOffState.eFault :
        bOut := FALSE;                                          // 故障态输出低 / output is low in the fault state
        IF rtReset.Q THEN
            eState := E_DL_MinOnOffState.eIdle;                 // 复位沿退出故障 / the reset edge leaves the fault state
        END_IF

ELSE
    // 强制安全兜底：非法状态一律回安全态并置故障（红线 R6）/ forced safe fallback for an illegal state
    eState := E_DL_MinOnOffState.eFault;                        // 强制回故障态 / force the fault state
    eErr   := 16#0001_039A;                                     // 非法状态（故障级）/ illegal state, fault level
    bError := TRUE;                                             // 置故障标志 / raise the fault flag
    bOut   := FALSE;                                            // 输出回安全态 / drive the output low
END_CASE

// 段 5｜守卫观测输出（只读定时器 ET，不做转移判据）/ segment 5, observable guard outputs, the elapsed time is never a transition test
bHoldOn  := (eState = E_DL_MinOnOffState.eHolding);              // 仅在保持态才算「强制延长运行」/ only the holding state really extends the run time
bHoldOff := (eState = E_DL_MinOnOffState.eCooldown);             // 冷却态即「强制延长停止」/ cooling down means the stop time is being enforced
IF (eState = E_DL_MinOnOffState.eStarting) OR (eState = E_DL_MinOnOffState.eHolding) THEN
    IF fbMinOn.ET < tMinOnEff THEN
        tRemaining := tMinOnEff - fbMinOn.ET;                    // 最短运行剩余 / remaining minimum on time
    ELSE
        tRemaining := DL_TIME_ZERO;                              // 已满 / already satisfied
    END_IF
ELSIF eState = E_DL_MinOnOffState.eCooldown THEN
    IF fbMinOff.ET < tMinOffEff THEN
        tRemaining := tMinOffEff - fbMinOff.ET;                  // 最短停止剩余 / remaining minimum off time
    ELSE
        tRemaining := DL_TIME_ZERO;                              // 已满 / already satisfied
    END_IF
ELSE
    tRemaining := DL_TIME_ZERO;                                  // 无守卫 / no guard active
END_IF
END_FUNCTION_BLOCK

(* ---- FB_DL_MinPulseWidthFilter.st ---- *)
(*==============================================================================
 * 组件名称 (Component)  : FB_DL_MinPulseWidthFilter
 * 溯源说明 (Provenance) : IEC 61131-3 标准语义的道莅防御性实现（零检索变体线）
 * 所属子库 (Sublibrary) : DL_Base / SignalShape
 * 当前版本 (Version)    : 1.0.0
 * 兼容性   (Platform)   : CODESYS 3.5 / TwinCAT 3 / 汇川 InoProShop；
 *                         纯 IEC 61131-3（第 3 版），仅用标准库 TON
 * 组件分类 (Category)   : 功能块（TYPE E_DL_MinPulseState :
(
    ePassThrough := 0, // 直通模式：双零参数 / Pass-through: both widths zero
    eStableLow   := 1, // 稳态低：等待有效接通 / Stable low: waiting qualified on
    eStableHigh  := 2  // 稳态高：等待有效断开 / Stable high: waiting qualified off
);
END_TYPE

FUNCTION_BLOCK）· 最小脉宽滤波
 * 功能一句话 (Summary)  : 抑制窄于 tMinOn / tMinOff 的毛刺，达标脉冲 1:1 透传。
 * 边界与安全 (Boundary) : ①两相超时参数为负 → 钳 0 并置故障码 0001_03BF；
 *                         ②两参数同为 0 → 直通模式（边沿即透传）；
 *                         ③上电输出初始化 FALSE，首扫无假触发；
 *                         ④两相定时器无条件周期刷新，不包 IF 跳调。
 * 错误码    : 16#0001_03BF 两相超时参数非法（负值已钳 0）——故障级
 *             16#0001_03C0 保留禁用（不得挪用，本件零赋值）
 * 码位总账  : 16#0001_03BF 用 ｜ 16#0001_03C0 预留
 * 修改记录  : v1.0.0 R26 初版
 *==============================================================================*)
FUNCTION_BLOCK FB_DL_MinPulseWidthFilter
VAR_INPUT
    bIn      : BOOL; // 待滤波信号输入 / Signal to be filtered
    tMinOn   : TIME; // 最小接通脉宽 [ms] / Minimum on-pulse width [ms]
    tMinOff  : TIME; // 最小断开脉宽 [ms] / Minimum off-pulse width [ms]
END_VAR
VAR_OUTPUT
    bOut        : BOOL; // 滤波后输出，达标脉冲 1:1 透传 / Filtered output, qualified pulses pass 1:1
    bSuppressed : BOOL; // 本周期有脉冲被抑制标志 / A glitch is being suppressed this cycle
    eErr        : UDINT; // 本周期错误码，0=无错 / Error code this cycle, 0 = none
END_VAR
VAR
    eState  : E_DL_MinPulseState; // 两相滤波状态机当前态 / Two-phase filter state machine state
    bOutIni : BOOL; // 输出初始化哨兵，恒 FALSE 保证上电安全侧 / Output init sentinel, stays FALSE for safe power-up
    tonOn   : TON; // 接通保持计时，验证接通脉宽达标 / On-hold timer, validates on-pulse width
    tonOff  : TON; // 断开保持计时，验证断开脉宽达标 / Off-hold timer, validates off-pulse width
    tOnEff  : TIME; // 接通脉宽有效值（钳位后）/ Effective on-width after clamping
    tOffEff : TIME; // 断开脉宽有效值（钳位后）/ Effective off-width after clamping
END_VAR
VAR CONSTANT
    cTZero : TIME := T#0MS; // 零时长基准 / Zero-duration baseline
END_VAR

// ---------- 两相定时器无条件周期刷新（不包 IF，防漏调） ----------
tonOn (IN := (bIn) AND (eState = E_DL_MinPulseState.eStableLow),  PT := tOnEff);
tonOff(IN := (NOT bIn) AND (eState = E_DL_MinPulseState.eStableHigh), PT := tOffEff);

// ---------- 参数防御：负值钳 0 并置码；双零转直通 ----------
eErr := 0;
IF (TIME_TO_DINT(tMinOn) < 0) OR (TIME_TO_DINT(tMinOff) < 0) THEN
    tOnEff  := cTZero;                       // 负值钳 0 / Clamp negative to zero
    tOffEff := cTZero;
    eErr    := 16#0001_03BF;                 // 故障级：参数非法已钳 / fault: illegal params clamped
ELSIF (tMinOn = cTZero) AND (tMinOff = cTZero) THEN
    tOnEff  := cTZero;                       // 直通模式配置 / Pass-through configuration
    tOffEff := cTZero;
ELSE
    tOnEff  := tMinOn;                       // 参数合法原样采用 / Legal params used as-is
    tOffEff := tMinOff;
END_IF

// ---------- 两相状态机：稳态低等待有效接通，稳态高等待有效断开 ----------
CASE eState OF
    E_DL_MinPulseState.ePassThrough:
        bOut := bIn;                          // 双零直通，边沿即透传 / Pass-through, edges pass at once

    E_DL_MinPulseState.eStableLow:            // 拍 N 进入：输出保持低 / Entered: output held low
        bOut := FALSE;                        // 本拍行为：未达标脉冲被吸收 / This cycle: short pulses absorbed
        IF tonOn.Q THEN                       // 接通保持达标（定时器含 bIn 条件，Q 为真即 bIn 持续达标）
            bOut    := TRUE;                  // 转出：输出抬升 / Leaving: output rises
            eState  := E_DL_MinPulseState.eStableHigh;
        END_IF

    E_DL_MinPulseState.eStableHigh:           // 拍 N 进入：输出保持高 / Entered: output held high
        bOut := TRUE;                         // 本拍行为：达标脉冲透传 / This cycle: qualified pulse passes
        IF tonOff.Q THEN                      // 断开保持达标 / Off-hold qualified
            bOut    := FALSE;                 // 转出：输出回落 / Leaving: output falls
            eState  := E_DL_MinPulseState.eStableLow;
        END_IF

    ELSE                                      // 非法状态兜底，归安全态低电平 / Illegal state fallback to safe low
        eState := E_DL_MinPulseState.eStableLow;
        bOut   := FALSE;
END_CASE

// ---------- 抑制标志：输入与输出不一致即处于毛刺吸收期 ----------
IF bIn <> bOut THEN
    bSuppressed := TRUE;                      // 毛刺吸收中 / Glitch being absorbed
ELSE
    bSuppressed := FALSE;                     // 同拍清除，无生命周期残留 / Same-cycle clear, no latch residue
END_IF

END_FUNCTION_BLOCK

(* ---- FB_DL_ModeArbiter.st ---- *)
(*==============================================================================
 * 组件名称 (Component)  : FB_DL_ModeArbiter
 * 所属子库 (Sublibrary) : DL_Base
 * 当前版本 (Version)    : 1.0.0
 * 兼容性   (Platform)   : CODESYS 3.5+ / TwinCAT 3 / 汇川 InoProShop / 施耐德 Machine Expert
 *                         仅依赖 Standard.library（R_TRIG），零厂商私有库
 * 功能描述 (Function)   : 三源运行模式请求仲裁：手动（Manual）> 自动（Auto）> 远程（Remote）
 *                         三级优先。请求为电平输入，模式**进入**必须由对应请求的上升沿
 *                         （或 bActManual 手动激活沿）触发；高优先级请求沿出现即抢占当前
 *                         低级模式（bPreempted 记录被顶事实）；高优先级撤销后**不自动回退**
 *                         到低级模式——回退必须由低级请求重新沿触发，防模式振荡；全部请求
 *                         撤销 → eNone（不记忆最后模式，HMI 记忆语义由上层做）。
 *                         多请求同拍 → 按优先级电平取最高级裁决，同拍置 bChanged。
 * 接口     (Interface)  : 输入 bReqManual / bReqAuto / bReqRemote 三源请求电平、
 *                         bActManual 手动激活沿源（如本地选择开关）；输出 eMode 当前模式、
 *                         bChanged 模式变更单拍、bPreempted 被抢占单拍。
 * 边界     (Boundary)   : ① **属主边界（写死）：本件只做模式请求仲裁与状态出口，不驱动任何
 *                         执行器、不做模式内的动作编排**；模式内行为由上层按 eMode 分发。
 *                         ② 进入 eManual 的沿条件 = rtReqManual 上升沿 ∨ (bActManual 上升沿
 *                         ∧ bReqManual 电平为真)；bActManual 单独出现而手动请求电平不成立时
 *                         不进入手动模式（防无保持电平的闪进闪出）。
 *                         ③ 在模式中保持条件 = 本模式请求电平为真；电平撤销即回 eNone，
 *                         **不**顺延到仍为真的低级请求（不自动回退铁律，回退必须重新沿触发）。
 *                         ④ 抢占定义：在非 eNone 模式中，被更高优先级的请求沿（或手动激活沿）
 *                         顶出 → bPreempted 单拍 + bChanged 单拍；平级沿（本模式自身请求沿）
 *                         不算抢占、不算变更。
 *                         ⑤ bActManual 在自动/远程模式中同样具备抢占能力（手动永远最高优先），
 *                         前提仍是 bReqManual 电平为真。
 *                         ⑥ 零全局耦合（无 GVL / 无 VAR_EXTERNAL / 无物理地址）。
 * 分工声明 (Scope)      : 与 `FB_DL_MutexOwnerAudit` 分工：运行模式 ≠ 互斥锁属主，那件审计
 *                         资源占用属主，本件仲裁人机操作模式；与 `FB_DL_DeviceHealthArbiter`
 *                         分工：健康裁决域归那件，本件不读任何健康量。
 * 来源标签 (Source Tag) : 自研线（公开优先级仲裁语义 clean-room）
 * 码表     (Codes)      : 本件不占用任何全局数字码位。出口为 ENUM 模式 + BOOL 组；
 *                         数字码位待主控收口阶段统一派号。
 * 红线自检 (Redline)    : R1 ✓ 零 GVL/VAR_EXTERNAL ｜ R2 ✓ 零 %I/%Q/%M ｜ R3 ✓ 纯 IEC 61131-3
 *                         R4 N/A（无浮点运算） ｜ R5 ✓ 声明逐行同行双语注释
 *                         R6 ✓ ENUM+CASE 含 ELSE ｜ R7 ✓ 四 R_TRIG 段 0 无条件刷新
 * 修订历史 (Revision)   : 2026-11-20  v1.0.0  R48 首版（批次 1 · 序号 4）
 *                         验收向量：手动沿抢占自动 → bPreempted；手动电平撤销 → eNone 不回
 *                         自动；自动沿重触发 → eAuto；三沿同拍 → eManual 优先。
 *==============================================================================*)

TYPE E_DL_MarMode :
(
    eNone   := 0,    // 无有效模式（全部请求撤销）/ No active mode
    eManual := 10,   // 手动模式（最高优先级）/ Manual mode, highest priority
    eAuto   := 20,   // 自动模式（中优先级）/ Auto mode, middle priority
    eRemote := 30    // 远程模式（最低优先级）/ Remote mode, lowest priority
);
END_TYPE

FUNCTION_BLOCK FB_DL_ModeArbiter
VAR_INPUT
    bReqManual : BOOL := FALSE;   // 手动模式请求电平 [-] / Manual mode request level
    bReqAuto   : BOOL := FALSE;   // 自动模式请求电平 [-] / Auto mode request level
    bReqRemote : BOOL := FALSE;   // 远程模式请求电平 [-] / Remote mode request level
    bActManual : BOOL := FALSE;   // 手动激活沿源（如本地选择开关动作；须伴随手动请求电平才生效） [-] / Manual activation edge source, needs manual request level
END_VAR
VAR_OUTPUT
    eMode      : E_DL_MarMode;    // 当前模式出口 [-] / Current mode outlet
    bChanged   : BOOL;            // 模式变更，单拍脉冲 [-] / Mode changed, single-scan pulse
    bPreempted : BOOL;            // 被高优先级抢占，单拍脉冲 [-] / Preempted by higher priority, single-scan pulse
END_VAR
VAR
    _eMode    : E_DL_MarMode := E_DL_MarMode.eNone;   // 内部模式（CASE 唯一写入目标） / Internal mode
    rtReqMan  : R_TRIG;           // 手动请求沿实例，段 0 无条件调用 / Manual request edge instance
    rtReqAuto : R_TRIG;           // 自动请求沿实例，段 0 无条件调用 / Auto request edge instance
    rtReqRem  : R_TRIG;           // 远程请求沿实例，段 0 无条件调用 / Remote request edge instance
    rtActMan  : R_TRIG;           // 手动激活沿实例，段 0 无条件调用 / Manual activation edge instance
    _bChanged : BOOL;             // 变更单拍内部量（统一出口映射，R34 两段式） / Changed pulse internal
    _bPreempt : BOOL;             // 抢占单拍内部量（统一出口映射） / Preempted pulse internal
END_VAR

(* —— 段 0：四枚沿实例无条件周期刷新 —— *)
rtReqMan(CLK := bReqManual);    // 手动请求沿，每拍必调 / Manual request edge, every scan
rtReqAuto(CLK := bReqAuto);     // 自动请求沿，每拍必调 / Auto request edge, every scan
rtReqRem(CLK := bReqRemote);    // 远程请求沿，每拍必调 / Remote request edge, every scan
rtActMan(CLK := bActManual);    // 手动激活沿，每拍必调 / Manual activation edge, every scan

(* —— 段 1：单拍量预清零（_eMode 为锁存状态量不入清单，R107） —— *)
bChanged   := FALSE;            // 变更脉冲预清 / Changed pulse preset
bPreempted := FALSE;            // 抢占脉冲预清 / Preempted pulse preset
_bChanged  := FALSE;            // 内部变更脉冲预清 / Internal changed pulse preset
_bPreempt  := FALSE;            // 内部抢占脉冲预清 / Internal preempted pulse preset

(* —— 段 2：模式状态机（进入必沿触发、保持必电平、撤销不回退） —— *)
CASE _eMode OF

E_DL_MarMode.eNone:
    IF rtReqMan.Q OR (rtActMan.Q AND bReqManual) THEN
        _eMode := E_DL_MarMode.eManual;                 // 手动沿（或激活沿∧手动电平）入手动 / Manual edge enters manual
        _bChanged := TRUE;                              // 记变更 / Mark changed
    ELSIF rtReqAuto.Q THEN
        _eMode := E_DL_MarMode.eAuto;                   // 自动沿入自动 / Auto edge enters auto
        _bChanged := TRUE;                              // 记变更 / Mark changed
    ELSIF rtReqRem.Q THEN
        _eMode := E_DL_MarMode.eRemote;                 // 远程沿入远程 / Remote edge enters remote
        _bChanged := TRUE;                              // 记变更 / Mark changed
    END_IF                                              // 同拍多沿按优先级顺序裁决（IF-ELSIF 级联即优先级）/ Same-scan multi-edge resolved by priority cascade

E_DL_MarMode.eManual:
    IF NOT bReqManual THEN
        _eMode := E_DL_MarMode.eNone;                   // 手动电平撤销 → eNone，不自动回退（铁律③）/ Manual level dropped, no auto fallback
        _bChanged := TRUE;                              // 记变更 / Mark changed
    ELSIF rtReqAuto.Q THEN
        _eMode := E_DL_MarMode.eAuto;                   // 自动沿抢占手动 / Auto edge preempts manual
        _bPreempt := TRUE;                              // 记抢占 / Mark preempted
        _bChanged := TRUE;                              // 记变更 / Mark changed
    ELSIF rtReqRem.Q THEN
        _eMode := E_DL_MarMode.eRemote;                 // 远程沿抢占手动 / Remote edge preempts manual
        _bPreempt := TRUE;                              // 记抢占 / Mark preempted
        _bChanged := TRUE;                              // 记变更 / Mark changed
    END_IF

E_DL_MarMode.eAuto:
    IF NOT bReqAuto THEN
        _eMode := E_DL_MarMode.eNone;                   // 自动电平撤销 → eNone，不自动回退 / Auto level dropped, no auto fallback
        _bChanged := TRUE;                              // 记变更 / Mark changed
    ELSIF rtReqMan.Q OR (rtActMan.Q AND bReqManual) THEN
        _eMode := E_DL_MarMode.eManual;                 // 手动沿抢占自动 / Manual edge preempts auto
        _bPreempt := TRUE;                              // 记抢占 / Mark preempted
        _bChanged := TRUE;                              // 记变更 / Mark changed
    ELSIF rtReqRem.Q THEN
        _eMode := E_DL_MarMode.eRemote;                 // 远程沿抢占自动 / Remote edge preempts auto
        _bPreempt := TRUE;                              // 记抢占 / Mark preempted
        _bChanged := TRUE;                              // 记变更 / Mark changed
    END_IF

E_DL_MarMode.eRemote:
    IF NOT bReqRemote THEN
        _eMode := E_DL_MarMode.eNone;                   // 远程电平撤销 → eNone，不自动回退 / Remote level dropped, no auto fallback
        _bChanged := TRUE;                              // 记变更 / Mark changed
    ELSIF rtReqMan.Q OR (rtActMan.Q AND bReqManual) THEN
        _eMode := E_DL_MarMode.eManual;                 // 手动沿抢占远程 / Manual edge preempts remote
        _bPreempt := TRUE;                              // 记抢占 / Mark preempted
        _bChanged := TRUE;                              // 记变更 / Mark changed
    ELSIF rtReqAuto.Q THEN
        _eMode := E_DL_MarMode.eAuto;                   // 自动沿抢占远程 / Auto edge preempts remote
        _bPreempt := TRUE;                              // 记抢占 / Mark preempted
        _bChanged := TRUE;                              // 记变更 / Mark changed
    END_IF

ELSE
    _eMode := E_DL_MarMode.eNone;                       // 非法模式兜底拉回无模式 / Illegal mode falls back to none
    _bChanged := TRUE;                                  // 兜底迁移也记变更 / Fallback marks changed

END_CASE

(* —— 段 3：出口单点映射（bChanged/bPreempted 由内部量统一映射，R34 两段式；R191 同源） —— *)
bChanged   := _bChanged;                                // 变更单拍出口 / Changed pulse outlet
bPreempted := _bPreempt;                                // 抢占单拍出口 / Preempted pulse outlet
eMode      := _eMode;                                   // 当前模式出口 / Current mode outlet

END_FUNCTION_BLOCK

(* ---- FB_DL_ModuloCounter.st ---- *)
(*==============================================================================
 * 组件名称 (Component)  : FB_DL_ModuloCounter
 * 所属子库 (Sublibrary) : DL_Base
 * 当前版本 (Version)    : 1.0.0
 * 兼容性   (Platform)   : CODESYS 3.5 / TwinCAT 3 / 汇川 InoProShop / Machine Expert
 *                         仅依赖 Standard.library（R_TRIG），零厂商方言
 * 分类     (Category)   : 信号处理功能块（Function Block · 取模工位索引）
 * 功能简述 (Function)   : 循环计数器（转盘/弹夹工位索引）。0..(nMod-1) 取
 *                         模回绕，支持双向步进、带合法性校验的跳步与回绕事
 *                         件一拍输出；模数 <2 参数非法故障锁存，跳步目标越
 *                         界拒绝置信级，双向同拍抵消置信级。
 *                         与 FB_DL_EventCounter 职责分离（通用事件计数 vs
 *                         取模工位索引），非重复组件。
 * 公约遵循 (Convention) : 0.1/R23 事件型，免首扫——索引由步进/跳步沿驱动，
 *                         无初始化/跟踪同步语义，不设 bInit。
 *                         0.2/R21 bFault 为显式排除信息级码的派生式；信息级
 *                         只进 uErrorId 不进报警链。
 *                         0.7/R15 故障级锁存仅解除路径（bReset 上升沿）清码。
 *                         0.8 故障码段位 16#0001_xxxx（经 DL_Base VERSION.md
 *                         码表核对，0001_0103~0104 / 0001_0211 均未占用）：
 *                         【故障级】0001_0211 模数非法（nMod < 2）；
 *                         【信息级】0001_0103 跳步目标越界拒绝、0001_0104
 *                         双向步进同拍抵消。
 * 红线自检 (Redline)    : R1 零全局变量表/外部变量引用 ✓｜R2 零物理 IO 地址 ✓
 *                         R3 纯 IEC 61131-3 ✓｜R4 模数非法/越界防御 + 显式
 *                         类型转换（UINT↔DINT）✓
 *                         R5 全变量中英双语同行注释 ✓｜R7 边沿实例主体最前
 *                         部无条件刷新 ✓｜R8 常量化无魔法数 ✓
 * 设计要点 (Key notes)  : ① 取模实现禁用取余运算符对负数的平台差异——回绕
 *                           用条件加减法（减 nMod / 加 nMod）实现，全部在
 *                           DINT 域运算后显式转回 UINT（CODESYS/TwinCAT/
 *                           汇川三平台行为一致，跨平台意图注释在此留档）；
 *                         ② nMod < 2 → 参数非法故障锁存【故障级】（除零与
 *                           退化防御）；nJumpTo >= nMod → 跳步拒绝 + 信息级；
 *                         ③ bStepFwd 与 bStepRev 同拍到达：抵消，置信级；
 *                         ④ bWrapped 跨零点步进置位一拍（转盘单圈计数用）。
 * 开源溯源 (Origin)     : 来源标签 lgf-counter（RAW_NOTES_R7 S-1：LGF 库计
 *                         数器族的取模索引功能域语义，公开文档，仅借鉴功能
 *                         域；条件加减法回绕、跳步校验、故障码与引脚契约
 *                         100% 本库独立设计，clean-room 未复制源码）。
 * 验收向量 (Acceptance) :
 *   V1 连续步进跨零回绕：nMod=8，uIndex=7 时 bStepFwd → 0 且 bWrapped 一拍；
 *   V2 反向跨零：uIndex=0 时 bStepRev → 7 且 bWrapped 一拍；
 *   V3 合法跳步：nJumpTo=5 < nMod=8 → uIndex=5；非法跳步 nJumpTo=9 → 拒绝
 *      保持 5 且信息级 0001_0103；
 *   V4 模数=2 边界：uIndex 在 0/1 间循环；nMod=1 → 故障锁存 0001_0211；
 *   V5 双向抵消：同拍 bStepFwd+bStepRev → 不变且信息级 0001_0104；
 *   V6 复位：bReset 沿 → uIndex=0、故障清零。
 * 修订历史 (Revision)   :
 *   2026-11-15  v1.0.0  首版入库（Round 07 · DL_Base LGF Counter 组开组）
 *============================================================================*)
FUNCTION_BLOCK FB_DL_ModuloCounter
VAR_INPUT
    bStepFwd : BOOL;            // 前进步进脉冲（Step forward），R_TRIG 上升沿 +1 取模 / Step forward edge, +1 modulo
    bStepRev : BOOL;            // 后退步进脉冲（Step reverse），R_TRIG 上升沿 -1 取模 / Step reverse edge, -1 modulo
    bJump    : BOOL;            // 跳步指令（Jump to index），上升沿装载 nJumpTo（带合法性校验）/ Jump edge loads nJumpTo with validity check
    nJumpTo  : UINT;            // 跳步目标工位号（Jump target index）[-]，域 0..nMod-1，越界拒绝 / Jump target, range 0..nMod-1, rejected outside
    nMod     : UINT := 8;       // 循环模数（Modulo count，工位数）[-]，域 2..65535，禁止 0/1（除零与退化防御）/ Modulo count, range 2..65535, 0/1 forbidden
    bReset   : BOOL;            // 上升沿复位故障与清零（Reset edge clears fault and index）/ Rising edge resets fault and clears index
END_VAR
VAR_OUTPUT
    uIndex   : UINT;            // 当前工位索引（Current index）[-]，0..nMod-1 / Current station index, 0..nMod-1
    bWrapped : BOOL;            // 回绕事件标志（Wrapped event），跨零点步进置位一拍（转盘单圈计数用）/ Wrapped event, one scan when crossing zero point
    bFault   : BOOL;            // 故障标志（Fault flag），显式排除信息级码（R21）/ Fault flag, info codes explicitly excluded
    uErrorId : UDINT;           // 故障码（Error code），16#0001_xxxx 段，0=无故障 / Error code, family 16#0001_xxxx, 0 = none
END_VAR
VAR
    _fbTrigFwd   : R_TRIG;      // 前进沿检测（Forward edge detector）/ Forward step edge detector
    _fbTrigRev   : R_TRIG;      // 后退沿检测（Reverse edge detector）/ Reverse step edge detector
    _fbTrigJump  : R_TRIG;      // 跳步沿检测（Jump edge detector）/ Jump command edge detector
    _fbTrigReset : R_TRIG;      // 复位沿检测（Reset edge detector）/ Reset edge detector
    _bFaultLatch : BOOL;        // 故障锁存标志（Fault latch flag），仅 bReset 上升沿清除 / Fault latch, cleared only by reset edge
    _uErrorIdInt : UDINT;       // 内部故障级码寄存（Internal fault-level code register）/ Internal fault-level code register
    _uInfoCode   : UDINT;       // 本拍信息级码（Info code this cycle），瞬时型每拍重算 / Transient info code, recomputed each scan
    _bFwdEdge    : BOOL;        // 本拍前进沿有效（Forward edge active this scan）/ Forward edge this scan
    _bRevEdge    : BOOL;        // 本拍后退沿有效（Reverse edge active this scan）/ Reverse edge this scan
    _bJumpEdge   : BOOL;        // 本拍跳步沿有效（Jump edge active this scan）/ Jump edge this scan
    _nWork       : DINT;        // DINT 域索引工作副本（DINT-domain working index）[-]，条件加减法载体 / DINT working index for conditional wrap arithmetic
    _nModEff     : UINT := 8;   // 防御后生效模数（Sanitized effective modulo）[-] / Sanitized effective modulo
    _nModD       : DINT;        // 生效模数 DINT 镜像（DINT mirror of effective modulo）[-] / DINT mirror of the modulo
END_VAR

// ============================================================================
// 段 1｜边沿实例无条件周期刷新（R7/0.5：严禁置于 IF/CASE 分支内）
//      Unconditional per-cycle refresh of all edge instances (R7/0.5)
// ============================================================================
_fbTrigFwd(CLK   := bStepFwd);
_fbTrigRev(CLK   := bStepRev);
_fbTrigJump(CLK  := bJump);
_fbTrigReset(CLK := bReset);
_bFwdEdge  := _fbTrigFwd.Q;     // 本拍前进沿（Forward edge this scan）
_bRevEdge  := _fbTrigRev.Q;     // 本拍后退沿（Reverse edge this scan）
_bJumpEdge := _fbTrigJump.Q;    // 本拍跳步沿（Jump edge this scan）

// ============================================================================
// 段 2｜信息级码预清零 + 复位路径（R15：锁存型故障只在解除路径清码）
//      Info code preset zero + reset path (R15)
// ============================================================================
_uInfoCode := 0;                // 信息级瞬时型每拍重算（Transient info recomputed each scan）
bWrapped := FALSE;              // 回绕事件每拍预清零，由段 4 事件置位一拍（Wrapped flag preset FALSE, set one scan by stage 4）

IF _fbTrigReset.Q THEN
    uIndex      := 0;           // 索引清零（Index cleared）
    _bFaultLatch := FALSE;      // 故障锁存解除（Fault latch released）
    _uErrorIdInt := 16#0000_0000; // 故障码清零（Fault code cleared）
END_IF

// ============================================================================
// 段 3｜参数防御：nMod < 2 → 故障锁存（0/1 除零与退化防御，故障级）
//      Parameter guard: nMod < 2 latches a fault (divide-by-zero and degeneration)
// ============================================================================
IF nMod < 2 THEN
    _bFaultLatch := TRUE;              // 模数非法故障锁存（Invalid modulo latch）
    _uErrorIdInt := 16#0001_0211;      // 0001_0211 模数非法【故障级】/ Invalid modulo, fault level
ELSE
    _nModEff := nMod;                  // 生效模数镜像（Effective modulo mirror）
    _nModD   := UINT_TO_DINT(_nModEff); // 显式转换 DINT 域（Explicit conversion to DINT domain）

    // ========================================================================
    // 段 4｜索引主逻辑：双向抵消 → 跳步 → 单向步进（条件加减法回绕）
    //      Index main logic: dual cancellation, jump, then conditional wrap stepping
    // ========================================================================
    IF _bFwdEdge AND _bRevEdge THEN
        _uInfoCode := 16#0001_0104;    // 0001_0104 双向同拍抵消【信息级】，索引不变 / Dual steps cancel, index unchanged, info level
    ELSIF _bJumpEdge THEN
        IF nJumpTo < _nModEff THEN
            uIndex := nJumpTo;         // 合法跳步：目标域 0..nMod-1（Valid jump within domain）
        ELSE
            _uInfoCode := 16#0001_0103; // 0001_0103 跳步目标越界拒绝【信息级】，索引保持 / Jump target out of range, rejected, info level
        END_IF
    ELSIF _bFwdEdge OR _bRevEdge THEN
        _nWork := UINT_TO_DINT(uIndex); // 显式转换进 DINT 域运算（Explicit conversion into DINT arithmetic）
        IF _bFwdEdge THEN
            _nWork := _nWork + 1;      // 前进一步（Forward one step）
            IF _nWork >= _nModD THEN
                _nWork := 0;           // 条件加减法回绕：越过模数回零点（Conditional wrap: above modulo back to zero, no remainder operator）
                bWrapped := TRUE;      // 跨零点事件一拍（Wrapped event, one scan）
            END_IF
        ELSE
            _nWork := _nWork - 1;      // 后退一步（Reverse one step）
            IF _nWork < 0 THEN
                _nWork := _nModD - 1;  // 条件加减法回绕：越过零点回模数尾（Conditional wrap: below zero to modulo tail）
                bWrapped := TRUE;      // 跨零点事件一拍（Wrapped event, one scan）
            END_IF
        END_IF
        uIndex := DINT_TO_UINT(_nWork); // 显式转换回 UINT 单点出口（Explicit conversion back, single outlet）
    END_IF
END_IF

// ============================================================================
// 段 5｜bFault/uErrorId 出口（R21：bFault 显式排除信息级；无故障级锁存时
//       uErrorId 透出本拍信息级码）
//      Outlets: bFault excludes info codes (R21); uErrorId shows info code when no fault
// ============================================================================
bFault := _bFaultLatch;             // 故障级派生式（Fault-level derived form）
IF _bFaultLatch THEN
    uIndex := 0;                    // 故障期索引输出安全零（Safe zero while latched）
    uErrorId := _uErrorIdInt;       // 故障级码优先透出（Fault-level code has priority）
ELSE
    uErrorId := _uInfoCode;         // 无故障时透出本拍信息级码（Transient info code when no fault）
END_IF
END_FUNCTION_BLOCK

(* ---- FB_DL_MultiClickDetect.st ---- *)
(*
  FB_DL_MultiClickDetect  —  按钮短按/长按/双击三形态判定 / Button short, long and double-click detection
  分类 Category : DL_Base
  版本 Version  : 1.0.0
  来源 Source   : t1-5-tcopen — 调试盘人机交互族零检索深化
  溯源 Origin   : clean-room 实现，未复制任何源码行
  功能 Function : 1) 对 bBtn 判定三种按压形态：短按（释放早于 tLong 且无双击窗内第二沿）、
                  长按（按压持续达 tLong）、双击（释放后 tDouble 窗内出现第二按压沿）；
                  2) bShortPulse / bDouble 单拍脉冲在判定拍发出；bLong 在达窗拍发出单拍脉冲；
                  3) 双击窗内第二沿判据使用当拍量（rtPrs.Q），无锁存量自指；
                  4) bReset 上升沿清组态故障锁存。
  边界 Boundary : ① 组态闸：tLong > tDouble > T#0S 必须成立，违例置故障级 03DE，三脉冲出口强制 FALSE；
                  ② 长按期间释放不产生短按脉冲（长按优先归因，防同拍双归因）；
                  ③ 状态机 ENUM+CASE 全覆盖 + ELSE 兜底落 03DF 故障锁存；
                  ④ 无 GVL 依赖：纯引脚输入输出，无外部变量引用，无物理 IO 地址。
  依赖 Depends  : 仅 Standard.library（TON / R_TRIG）
  码表 Error codes（段 0001，窗口 03DE~03DF / 04A1~04A2）:
    16#0001_03DE 故障级：组态非法（tLong <= tDouble 或任一窗 <= T#0S），锁存至 bReset
    16#0001_03DF 故障级：状态机落 ELSE 兜底（非法相位 ID），锁存至 bReset
    16#0001_04A1 信息级：短按事件（与 bShortPulse 同拍）
    16#0001_04A2 信息级：双击事件（与 bDouble 同拍）
  修订历史 Revision :
    2026-11-19  v1.0.0  R41 首版（批次 1 · 序号 2）
*)

TYPE E_DL_McdState :
(
    eIdle   := 0,    // 空闲：按钮未按压 / Idle, button released
    eHeld   := 10,   // 按压中：等释放或达长按窗 / Held, waiting release or long window
    eWait2  := 20,   // 双击等待：释放早于长按窗，等第二沿 / Wait second press inside the double window
    eFault  := 90    // 故障：组态非法或兜底锁定 / Fault, latched
);
END_TYPE

FUNCTION_BLOCK FB_DL_MultiClickDetect
VAR_INPUT
    bBtn         : BOOL := FALSE;     // 按钮输入，TRUE = 按压 [-] / Button input, TRUE = pressed
    tLong        : TIME := T#1000MS;  // 长按窗 [ms]，必须 > tDouble / Long-press window
    tDouble      : TIME := T#300MS;   // 双击窗 [ms]，必须 > T#0S 且 < tLong / Double-click window
    bReset       : BOOL := FALSE;     // 复位，上升沿清故障锁存 / Reset edge clears fault latch
END_VAR
VAR_OUTPUT
    bShortPulse  : BOOL;              // 短按单拍脉冲 [-] / Short-press one-scan pulse
    bLong        : BOOL;              // 长按单拍脉冲 [-] / Long-press one-scan pulse
    bDouble      : BOOL;              // 双击单拍脉冲 [-] / Double-click one-scan pulse
    eState       : E_DL_McdState;     // 状态出口，段尾单点映射 / State outlet
    bError       : BOOL;              // 故障锁存标志 / Fault latch flag
    nErrId       : UDINT;             // 事件码，0 = 无事件 / Event code
END_VAR
VAR
    tonLongTo    : TON;               // 长按窗定时器（按压电平驱动），无条件刷新 / Long window timer
    tonDblTo     : TON;               // 双击窗定时器（等待相独占），无条件刷新 / Double window timer
    rtPrs        : R_TRIG;            // 按压沿实例，无条件刷新 / Press edge instance
    rtRel        : R_TRIG;            // 释放沿实例，无条件刷新 / Release edge instance
    rtReset      : R_TRIG;            // 复位沿实例，无条件刷新 / Reset edge instance
    _eState      : E_DL_McdState := E_DL_McdState.eIdle;  // 内部相位（CASE 唯一写入目标）/ Internal phase
    _uFault      : UDINT;             // 故障码锁存（锁存量）/ Latched fault code
    _uInfo       : UDINT;             // 信息码，每拍重算 / Transient info code
    _bLongSent   : BOOL;              // 本按压已发长按脉冲标志（防重复）/ Long pulse sent flag
    _bFault      : BOOL;              // 故障锁存位（锁存量）/ Latched fault bit
END_VAR

(* —— 段 0：定时器与沿实例无条件周期刷新（禁置于 IF/CASE 内） —— *)
rtPrs(CLK := bBtn);                       // 按压沿（每拍必调）
rtRel(CLK := NOT bBtn);                   // 释放沿（每拍必调）
rtReset(CLK := bReset);                   // 复位沿（每拍必调）
tonLongTo(IN := bBtn, PT := tLong);       // 长按窗（电平驱动，每拍必调）
tonDblTo(IN := (_eState = E_DL_McdState.eWait2), PT := tDouble);  // 双击窗（等待相独占，每拍必调）

(* —— 段 1：单拍量预清零（锁存量 _uFault/_bFault 不入清单；完成脉冲两段式出口） —— *)
_uInfo := 16#0000_0000;             // 信息码每拍重算
bShortPulse := FALSE;               // 短按脉冲缺省 FALSE
bLong := FALSE;                     // 长按脉冲缺省 FALSE
bDouble := FALSE;                   // 双击脉冲缺省 FALSE
nErrId := 16#0000_0000;             // 事件码缺省无事件

(* —— 段 2：复位沿与组态域闸（全当拍量判据） —— *)
IF rtReset.Q THEN                   // rtReset.Q = 当拍量
    _bFault := FALSE;               // 清故障锁存位
    _uFault := 16#0000_0000;        // 清故障锁存码
END_IF
IF (TIME_TO_DINT(tLong) <= TIME_TO_DINT(tDouble)) OR (TIME_TO_DINT(tDouble) <= 0) THEN
    _uFault := 16#0001_03DE;        // 故障级：组态非法
    _bFault := TRUE;
    _eState := E_DL_McdState.eIdle; // 故障期间回空闲
END_IF

(* —— 段 3：相位机（只判形态与发标志；脉冲在段 5 统一出口映射） —— *)
CASE _eState OF

E_DL_McdState.eIdle:
    IF rtPrs.Q AND (NOT _bFault) THEN
        _bLongSent := FALSE;            // 本按压长按脉冲未发
        _eState := E_DL_McdState.eHeld; // 进按压相
    END_IF

E_DL_McdState.eHeld:
    IF _bFault THEN
        _eState := E_DL_McdState.eIdle; // 故障相回空闲（脉冲出口已被强制 FALSE）
    ELSIF tonLongTo.Q AND (NOT _bLongSent) THEN
        bLong := TRUE;                  // 长按脉冲（本拍置位，段 5 出口同拍映射）
        _bLongSent := TRUE;             // 单发标志
    ELSIF rtRel.Q THEN
        IF (NOT _bLongSent) AND (TIME_TO_DINT(tDouble) > 0) THEN
            _eState := E_DL_McdState.eWait2;    // 早于长按窗释放：进双击等待相
        ELSE
            _eState := E_DL_McdState.eIdle;     // 长按后释放或组态异常：回空闲
        END_IF
    END_IF

E_DL_McdState.eWait2:
    IF _bFault THEN
        _eState := E_DL_McdState.eIdle;     // 故障相回空闲
    ELSIF rtPrs.Q THEN
        bDouble := TRUE;                    // 双击命中（窗内第二沿，当拍量判据）
        _uInfo := 16#0001_04A2;             // 信息级：双击事件
        _eState := E_DL_McdState.eHeld;     // 第二次按压继续按普通按压相处理
        _bLongSent := FALSE;                // 新按压重新计时长按
    ELSIF tonDblTo.Q THEN
        bShortPulse := TRUE;                // 双击窗超时：第一次按压判短按
        _uInfo := 16#0001_04A1;             // 信息级：短按事件
        _eState := E_DL_McdState.eIdle;     // 回空闲
    END_IF

E_DL_McdState.eFault:
    IF NOT _bFault THEN
        _eState := E_DL_McdState.eIdle;     // 故障解除（复位沿）回空闲，迁出边可达
    END_IF

ELSE
    _uFault := 16#0001_03DF;            // 故障级：非法相位 ID 兜底
    _bFault := TRUE;
    _eState := E_DL_McdState.eFault;    // 强制回故障相

END_CASE

(* —— 段 4：故障相脉冲出口强制 FALSE（安全侧，防故障期误发脉冲） —— *)
IF _bFault THEN
    bShortPulse := FALSE;           // 安全侧清脉冲
    bLong := FALSE;                 // 安全侧清脉冲
    bDouble := FALSE;               // 安全侧清脉冲
END_IF

(* —— 段 5：出口单点映射（锁存码回放，禁同拍抹除） —— *)
IF _bFault THEN
    nErrId := _uFault;              // 故障锁存码回放
ELSE
    nErrId := _uInfo;               // 信息码
END_IF
bError := _bFault;                  // 故障标志与锁存位同源
eState := _eState;                  // 状态出口单点映射

END_FUNCTION_BLOCK

(* ---- FB_DL_MultiSegmentTimer.st ---- *)
(*
  ==================================================================
  组件名 Component  : FB_DL_MultiSegmentTimer
  分类   Category   : DL_Base
  复杂度 Complexity  : 中
  版本   Version    : 1.0.0
  功能   Purpose    : 多段定时窗口组（日历窗）。8 段独立使能的日内分钟窗
                      （起止 0..1439），输出当前是否处于任一窗内 bInWindow、
                      当前活动段索引 nActiveSeg（-1 = 无）、段间重叠检测
                      bOverlap（信息级）与组态非法 bCfgErr。LGF Date and
                      Timer 多段定时语义 clean-room。
  来源   Source     : T2-1-lgf-date-timer（LGF 多段定时语义）
  溯源   Origin     : 日历窗多段定时为公开工程语义，clean-room 自研实现，
                      未复制 LGF 或任何厂商私有库源码。
  平台   Platform   : 纯 IEC 61131-3，CODESYS / TwinCAT / InoProShop 通用
  分工声明 Split     : 与 FB_DL_SchedWeekPlan 分工——后者做周计划调度，
                      本件做单日多段窗判定（无状态纯判定）。
  作者   Author     : 道莅代码库 · PLC 编程专家（R59）
  ------------------------------------------------------------------
  边界 Boundary     :
                      一 窗语义：[aStart, aStop) 左闭右开；aStart = aStop 视
                         为全日窗（1440 分钟）；支持 aStart > aStop 跨零点窗；
                      二 输入域闸：nNowMin ∉ [0..1439] 或任一使能段起止越域
                         → bCfgErr 置位，bInWindow 安全侧 FALSE（安全侧赋值
                         不受判定量污染）；
                      三 bOverlap 为信息级提示不锁存，不参与 bInWindow 判定；
                      四 无定时器无沿检测（无状态判定件），无全局变量、无
                         外部变量声明、无物理地址寻址。
  修订记录 Revision  :
    2026-11-21  v1.0.0  R59 首版（批 1 · 序号 3）
  ==================================================================
*)

FUNCTION_BLOCK FB_DL_MultiSegmentTimer
VAR_INPUT
    nNowMin : DINT;                     // 当日时刻 [分钟]，域 0..1439 / the minute of day, zero through one thousand four hundred thirty nine
    aEn     : ARRAY[0..7] OF BOOL;      // 段使能组（8 段独立使能）[-] / the segment enable array, eight independent enables
    aStart  : ARRAY[0..7] OF DINT;      // 段起始分钟组 [分钟]，域 0..1439 / the segment start minutes array
    aStop   : ARRAY[0..7] OF DINT;      // 段结束分钟组 [分钟]，域 0..1439 / the segment stop minutes array
END_VAR
VAR_OUTPUT
    bInWindow  : BOOL := FALSE; // 当前时刻处于任一使能窗内 [-] / the now inside any enabled window flag
    nActiveSeg : DINT := -1;    // 当前活动段索引，-1 = 无活动段 [段] / the active segment index, minus one when none
    bOverlap   : BOOL := FALSE; // 使能段间存在重叠（信息级）[-] / any enabled segments overlap, informational
    bCfgErr    : BOOL := FALSE; // 组态非法（时刻越域或使能段起止越域）[-] / the configuration fault
END_VAR
VAR CONSTANT
    DL_MST_SEGMAX : DINT := 8;    // 段容量上界 [段] / the segment capacity bound
    DL_MST_DAYMIN : DINT := 1440; // 全日分钟数 [分钟] / the minutes per day
END_VAR
VAR
    _nI    : DINT; // 段遍历索引（段判定环）/ the segment loop index
    _nJ    : DINT; // 重叠比对索引（重叠检测环）/ the overlap compare index
    _bHit  : BOOL; // 段命中工作量 [-] / the segment hit work flag
    _nSeg  : DINT; // 活动段寄存（-1 起步）/ the active segment register
    _bCfg  : BOOL; // 组态非法工作量（先算后出，避免多点回夹）/ the config fault work flag
    _bOvl  : BOOL; // 重叠工作量 / the overlap work flag
END_VAR

// 段 1｜输出预置与时刻域闸（安全侧赋值不受判定量污染，边界二）/ segment 1, the preset and the time domain gate
_bCfg := FALSE; // 组态非法工作量清零 / clear the config work flag
_bOvl := FALSE; // 重叠工作量清零 / clear the overlap work flag
_nSeg := -1; // 活动段预置无 / preset the active segment none
IF (nNowMin < 0) OR (nNowMin >= DL_MST_DAYMIN) THEN // 时刻越域 / the time out of domain
    _bCfg := TRUE; // 组态非法 / raise the config fault
END_IF

// 段 2｜使能段起止域校验与活动窗判定（含跨零点窗与全日窗语义，边界一）/ segment 2, the segment validation and the active window
FOR _nI := 0 TO DL_MST_SEGMAX - 1 DO // 逐段判定 / per segment verdict
    IF aEn[_nI] THEN // 段使能才校验与判定 / validate and judge only the enabled segment
        IF (aStart[_nI] < 0) OR (aStart[_nI] >= DL_MST_DAYMIN)
        OR (aStop[_nI] < 0) OR (aStop[_nI] >= DL_MST_DAYMIN) THEN // 起止越域 / the bounds out of domain
            _bCfg := TRUE; // 组态非法 / raise the config fault
        END_IF
        IF aStart[_nI] = aStop[_nI] THEN // 全日窗语义 / the full day window
            _bHit := TRUE; // 全日窗恒命中（越域统一由出口闸拦截）/ the full day window always hits
        ELSIF aStart[_nI] < aStop[_nI] THEN // 同日窗 [start, stop) / the same day window
            _bHit := (nNowMin >= aStart[_nI]) AND (nNowMin < aStop[_nI]); // 左闭右开命中 / the half open hit
        ELSE // 跨零点窗 [start, 1439] ∪ [0, stop) / the midnight spanning window
            _bHit := (nNowMin >= aStart[_nI]) OR (nNowMin < aStop[_nI]); // 双半区命中 / the two half zone hit
        END_IF
        IF _bHit AND (_nSeg < 0) THEN // 首个命中段为准（段号小者优先）/ the first hit segment wins
            _nSeg := _nI; // 记活动段 / register the active segment
        END_IF
    END_IF
END_FOR

// 段 3｜使能段两两重叠检测（信息级，边界三）/ segment 3, the pairwise overlap detection, informational
FOR _nI := 0 TO DL_MST_SEGMAX - 2 DO // 前段遍历 / the former loop
    IF aEn[_nI] AND (aStart[_nI] >= 0) AND (aStart[_nI] < DL_MST_DAYMIN)
    AND (aStop[_nI] >= 0) AND (aStop[_nI] < DL_MST_DAYMIN) THEN // 仅合法使能段参与比对 / only the valid enabled ones
        FOR _nJ := _nI + 1 TO DL_MST_SEGMAX - 1 DO // 后段遍历 / the latter loop
            IF aEn[_nJ] AND (aStart[_nJ] >= 0) AND (aStart[_nJ] < DL_MST_DAYMIN)
            AND (aStop[_nJ] >= 0) AND (aStop[_nJ] < DL_MST_DAYMIN) THEN // 仅合法使能段参与比对 / only the valid ones
                IF (aStart[_nI] < aStop[_nJ]) AND (aStart[_nJ] < aStop[_nI]) THEN // 区间相交判据（半开域交叠）/ the interval intersection
                    _bOvl := TRUE; // 置重叠提示 / raise the overlap hint
                END_IF
            END_IF
        END_FOR
    END_IF
END_FOR

// 段 4｜统一出口（安全侧：组态非法时 bInWindow 强制 FALSE，单点赋值）/ segment 4, the unified outlet
bCfgErr := _bCfg; // 组态非法出口 / the config fault outlet
bOverlap := _bOvl; // 重叠提示出口 / the overlap outlet
nActiveSeg := _nSeg; // 活动段出口 / the active segment outlet
IF _bCfg THEN // 组态非法安全侧 / the config fault safe side
    bInWindow := FALSE; // 窗内标志强制假 / force the window flag false
ELSE // 组态合法 / the valid configuration
    bInWindow := (_nSeg >= 0); // 命中即窗内 / the hit verdict
END_IF
END_FUNCTION_BLOCK
